(* Logix 5000 project; controller TFF vendor 1 type 14 code 107 rev 33.11; software revision 33.04; part 20 of 38 *)
(* tags used below, declared in another part *)
   Address : DINT;   // Temp Address
   Config : Configuration;   // Index Array used in configuration routines
   Index : DINT;   // Index
   TIME : DINT[2];
   TimeInSecondsDINT : DINT;
   AA008 : ALIAS FOR DigitalPoint[18];
   AI101 : ALIAS FOR AnalogPoint[16];
   AI101_SIG : ALIAS FOR DigitalPoint[106];
   AI104 : ALIAS FOR AnalogPoint[17];
   AI104_SIG : ALIAS FOR DigitalPoint[107];
   AI201A : ALIAS FOR AnalogPoint[10];
   AI201A_SIG : ALIAS FOR DigitalPoint[90];
   AI201B : ALIAS FOR AnalogPoint[0];
   AI201B_SIG : ALIAS FOR DigitalPoint[109];
   AI202 : ALIAS FOR AnalogPoint[9];
   AI202_SIG : ALIAS FOR DigitalPoint[105];
   AI203 : ALIAS FOR AnalogPoint[11];
   AI203_SIG : ALIAS FOR DigitalPoint[91];
   AI204 : ALIAS FOR AnalogPoint[12];
   AI204_SIG : ALIAS FOR DigitalPoint[92];
   AlarmAnalog : AlarmAnalog[50];   // Analog Alarm Array
   AlarmControl : AlarmControl;   // Alarm Control
   AlarmDeviation : AlarmDeviation[20];   // Control Loop Deviation Alarm Array
   AnalogOutput : AnalogOutput[25];   // Analog Output Array
   AnalogPoint : AnalogInput[50];   // Analog Input Array
   ARC_AI101 : ARC_pH;
   ARC_AI202 : ARC_pH;
   Concentration : Concentration;
   ControlLoop : ControlLoop[20];   // Control Loop Array
   ControlLoop_FeedBagLevel : ALIAS FOR ControlLoop[2];
   DF24VDC : ALIAS FOR DigitalPoint[4];
   DF24VDCPC : ALIAS FOR DigitalPoint[25];
   DF3PHP003 : ALIAS FOR DigitalPoint[27];
   DF48MIX : ALIAS FOR DigitalPoint[26];
   DF48P001 : ALIAS FOR DigitalPoint[23];
   DF48P002 : ALIAS FOR DigitalPoint[24];
   Diafiltration : Diafiltration;
   DigitalOutput : BOOL[256];   // Digital Output Array these bits are sent to output cards.
   DP : ALIAS FOR AnalogPoint[40];
   ES001 : ALIAS FOR DigitalPoint[2];
   ExternalTCU : BOOL;   // Use of External TCU
   ExternalWeight : BOOL;   // Use of External Weight
   FI003 : ALIAS FOR AnalogPoint[42];
   FI101 : ALIAS FOR AnalogPoint[19];
   FI101_SIG : ALIAS FOR DigitalPoint[110];
   FI201 : ALIAS FOR AnalogPoint[2];
   FI201_SIG : ALIAS FOR DigitalPoint[93];
   FI401 : ALIAS FOR AnalogPoint[20];
   FI401_SIG : ALIAS FOR DigitalPoint[94];
   LI101 : ALIAS FOR AnalogPoint[44];
   LI101Alarm : ALIAS FOR AlarmAnalog[44];
   MIX101 : ALIAS FOR AnalogPoint[14];
   MIX101_SIG : ALIAS FOR DigitalPoint[104];
   MIX101DF : ALIAS FOR DigitalPoint[28];
   Mixer : Mixer;   // Mixer config. structure
   NWP : ALIAS FOR AnalogPoint[45];
   Options : Options;   // Options List
   PCV101 : ALIAS FOR AnalogPoint[3];
   PCV101_Control : PCV_Control;   // PCV101 Control UDT
   PCV101_SIG : ALIAS FOR DigitalPoint[102];
   PCV201 : ALIAS FOR AnalogPoint[4];
   PCV201_Control : PCV_Control;   // PCV201 Control UDT
   PCV201_SIG : ALIAS FOR DigitalPoint[103];
   PERM : ALIAS FOR AnalogPoint[46];
   PI001 : ALIAS FOR AnalogPoint[5];
   PI001_SIG : ALIAS FOR DigitalPoint[97];
   PI101 : ALIAS FOR AnalogPoint[6];
   PI101_SIG : ALIAS FOR DigitalPoint[98];
   PI201 : ALIAS FOR AnalogPoint[7];
   PI201_SIG : ALIAS FOR DigitalPoint[99];
   PI401 : ALIAS FOR AnalogPoint[8];
   PI401_SIG : ALIAS FOR DigitalPoint[100];
   PI601 : ALIAS FOR AnalogPoint[21];
   PI601_SIG : ALIAS FOR DigitalPoint[95];
   PISL601 : ALIAS FOR DigitalPoint[0];
   PISL602 : ALIAS FOR DigitalPoint[1];
   PSH001 : ALIAS FOR DigitalPoint[21];
   PSH401 : ALIAS FOR DigitalPoint[22];
   SIC001 : ALIAS FOR Drive[1];
   SIC001DF : ALIAS FOR DigitalPoint[16];
   SIC002 : ALIAS FOR Drive[2];
   SIC002DF : ALIAS FOR DigitalPoint[17];
   SIC003DF : ALIAS FOR DigitalPoint[29];
   SIC004 : ALIAS FOR Drive[3];
   Tank : TankManagement;   // Tank Management
   TCU101 : ALIAS FOR AnalogPoint[18];
   TCU101_AO : ALIAS FOR AnalogOutput[6];
   TCU101_SIG : ALIAS FOR DigitalPoint[108];
   TCU101DF : ALIAS FOR DigitalPoint[30];
   TI101 : ALIAS FOR AnalogPoint[13];
   TI101_SIG : ALIAS FOR DigitalPoint[101];
   TI201 : ALIAS FOR AnalogPoint[22];
   TI201_SIG : ALIAS FOR DigitalPoint[111];
   TMP : ALIAS FOR AnalogPoint[41];
   Totalizer : Totalizers[20];   // Totalizers Array
   UserCr1 : ALIAS FOR DigitalPoint[65];
   UserCr2 : ALIAS FOR DigitalPoint[67];
   UserNCr1 : ALIAS FOR DigitalPoint[64];
   UserNCr2 : ALIAS FOR DigitalPoint[66];
   Valve : Valve[100];   // Valve Array
   WI101 : ALIAS FOR AnalogPoint[15];
   WI101Alarm : ALIAS FOR AlarmAnalog[15];
   WI201 : ALIAS FOR AnalogPoint[1];
   WI201_SIG : ALIAS FOR DigitalPoint[96];
   XV003 : ALIAS FOR Valve[2];
   XV004 : ALIAS FOR Valve[3];
   XV005 : ALIAS FOR Valve[4];
   XV006 : ALIAS FOR Valve[5];
   XV007 : ALIAS FOR Valve[6];
   YA01 : ALIAS FOR DigitalPoint[50];
   YA02 : ALIAS FOR DigitalPoint[51];
   YA03 : ALIAS FOR DigitalPoint[52];
   YA04 : ALIAS FOR DigitalPoint[53];
   YA05 : ALIAS FOR DigitalPoint[54];
   YA06 : ALIAS FOR DigitalPoint[55];
   YA07 : ALIAS FOR DigitalPoint[56];
   YA08 : ALIAS FOR DigitalPoint[57];
   YA09 : ALIAS FOR DigitalPoint[58];
   YA10 : ALIAS FOR DigitalPoint[59];
   YA11 : ALIAS FOR DigitalPoint[60];
   YA12 : ALIAS FOR DigitalPoint[61];
   YA13 : ALIAS FOR DigitalPoint[62];
   YA14 : ALIAS FOR DigitalPoint[63];
   YA15 : ALIAS FOR DigitalPoint[69];
   YA16 : ALIAS FOR DigitalPoint[70];
   YA17 : ALIAS FOR DigitalPoint[71];
   YA18 : ALIAS FOR DigitalPoint[72];
   YA41 : ALIAS FOR DigitalPoint[73];
   ZS008 : ALIAS FOR DigitalPoint[5];
   ZSDF : ALIAS FOR DigitalPoint[68];
(* Process, continued *)

ROUTINE Alarm_Init_Config   (* structured text *)
   (* =======================================================================
   	Alarm_Init_Config : initialize alarms to default values
   
   	List of treatments
   		- Analog alarms set point with scale Min and Max
   		- Deviation alarms
   		- Digital alarms
   	-----------------------------------------------------------------------------------------------------------------------------------------------------
   	History
   		2021-NOV-17 - Merck - Q.Spindler- Initial version for Candidate Release 1.01.00.00.a
   		2022-SEP-22 - Actemium - J. Jaekel - Modifications for Candidate Release 1.01.00.01.a
   			- Add TI201_SIG
   =============================================================================================================================*)
   
   (*Analog Set point to min/max scale, Enable alarm, timer to  2s
   ============================================================*)
   FOR Index := 0 to 49 by 1 do
   	IF AnalogPoint[Index].EnableCfg THEN
   		AlarmAnalog[Index].Override := 0; // Enable
   		AlarmAnalog[Index].LOLO := AnalogPoint[Index].ScaledMin ;
   		AlarmAnalog[Index].LO := AnalogPoint[Index].ScaledMin ;
   		AlarmAnalog[Index].HI := AnalogPoint[Index].ScaledMax ;
   		AlarmAnalog[Index].HIHI := AnalogPoint[Index].ScaledMax ;
   		AlarmAnalog[Index].LOLOTimerSP := 2 ;
   		AlarmAnalog[Index].LOTimerSP := 2 ;
   		AlarmAnalog[Index].HITimerSP := 2 ;
   		AlarmAnalog[Index].HIHITimerSP := 2 ;
   	END_IF;
   End_for ;
   
   (*Specific case for WI101
   ============================================================*)
   WI101Alarm.HI := Tank.Config.TankSelectPLC *1.2;
   WI101Alarm.HIHI := Tank.Config.TankSelectPLC *1.2;
   
   (*Specific case for LI101
   ============================================================*)
   LI101Alarm.HI := Tank.Config.TankSelectPLC;
   LI101Alarm.HIHI := Tank.Config.TankSelectPLC;
   
   (*Deviation alarm HI 100% HIHI 100%, Disable alarm, timer to 2s
   ============================================================*)
   FOR Index := 0 to 19 by 1 do
   	IF AlarmDeviation[Index].EnableCfg THEN
   		AlarmDeviation[Index].Override := 1; // Disable
   		AlarmDeviation[Index].HI := 100 ;
   		AlarmDeviation[Index].HIHI := 100 ;
   		AlarmDeviation[Index].HITimerSP := 2 ;
   		AlarmDeviation[Index].HIHITImerSP := 2 ;
   	END_IF;
   End_for ;
   
   (*Analog Set point to Disable alarm
   ============================================================*)
   // N/A
   
   (* Discrete Alarms
   ============================================================*)
   ES001.DelayTimerSP := 0;
   PISL601.Override := 0; PISL601.Priority := 1; PISL601.DelayTimerSP := 2;
   PISL602.Override := 0; PISL602.Priority := 1; PISL602.DelayTimerSP := 2;
   DF24VDC.Override := 0; DF24VDC.Priority := 1; DF24VDC.DelayTimerSP := 1;
   DF24VDCPC.Override := 0; DF24VDCPC.Priority := 1; DF24VDCPC.DelayTimerSP := 1;
   PSH001.Override := 0; PSH001.DelayTimerSP := 0;
   PSH401.Override := 0; PSH401.DelayTimerSP := 0;
   SIC001DF.Override := 0; SIC001DF.Priority := 1; SIC001DF.DelayTimerSP := 1;
   SIC002DF.Override := 0; SIC002DF.Priority := 1; SIC002DF.DelayTimerSP := 1;
   SIC003DF.Override := 0; SIC003DF.Priority := 1; SIC003DF.DelayTimerSP := 1;
   DF48P001.Override := 0; DF48P001.Priority := 1; DF48P001.DelayTimerSP := 1;
   DF48P002.Override := 0; DF48P002.Priority := 1; DF48P002.DelayTimerSP := 1;
   DF48MIX.Override := 0; DF48MIX.Priority := 1; DF48MIX.DelayTimerSP := 1;
   DF3PHP003.Override := 0; DF3PHP003.Priority := 1; DF3PHP003.DelayTimerSP := 1;
   AA008.Override := 0; AA008.Priority := 1; AA008.DelayTimerSP := 1;
   TCU101DF.Override := 0; TCU101DF.Priority := 1; TCU101DF.DelayTimerSP := 1;
   MIX101DF.Override := 0; MIX101DF.Priority := 1; MIX101DF.DelayTimerSP := 1;
   ZS008.Override := 0; ZS008.Priority := 1; ZS008.DelayTimerSP := 1;
   ZSDF.Override := 0; ZSDF.Priority := 1; ZSDF.DelayTimerSP := 1;
   
   
   YA01.Override := 0; YA01.Priority := 0; YA01.DelayTimerSP := 60;
   YA02.Override := 0; YA02.Priority := 0; YA02.DelayTimerSP := 60;
   YA03.Override := 0; YA03.Priority := 0; YA03.DelayTimerSP := 80;
   YA04.Override := 0; YA04.Priority := 0; YA04.DelayTimerSP := 60;
   YA05.Override := 0; YA05.Priority := 0; YA05.DelayTimerSP := 60;
   YA06.Override := 0; YA06.Priority := 1; YA06.DelayTimerSP := 5;
   YA07.Override := 0; YA07.Priority := 0; YA07.DelayTimerSP := 2;
   YA08.Override := 0; YA08.Priority := 1; YA08.DelayTimerSP := 5;
   YA09.Override := 0; YA09.Priority := 0; YA09.DelayTimerSP := 2;
   YA10.DelayTimerSP := 0;
   YA11.Override := 1; YA11.Priority := 0; YA11.DelayTimerSP := 5;
   YA12.Override := 0; YA12.Priority := 0; YA12.DelayTimerSP := 0;
   YA13.Override := 0; YA13.Priority := 0; YA13.DelayTimerSP := 2;
   YA14.Priority := 0; YA14.DelayTimerSP := 60;
   YA15.Override := 0; YA15.Priority := 1; YA15.DelayTimerSP := 5;
   YA16.Override := 1; YA16.Priority := 0; YA16.DelayTimerSP := 5;
   YA17.Override := 1; YA17.Priority := 0; YA17.DelayTimerSP := 5;
   YA18.Override := 0; YA18.Priority := 0; YA18.DelayTimerSP := 2;
   YA41.Override := 0; YA41.DelayTimerSP := 0;
   
   
   WI201_SIG.Override := 0; WI201_SIG.Priority := 0; WI201_SIG.DelayTimerSP := 10;
   MIX101_SIG.Override := 0; MIX101_SIG.Priority := 0; MIX101_SIG.DelayTimerSP := 10;
   AI101_SIG.Override := 0; AI101_SIG.Priority := 0; AI101_SIG.DelayTimerSP := 10;
   AI104_SIG.Override := 0; AI104_SIG.Priority := 0; AI104_SIG.DelayTimerSP := 10;
   TI101_SIG.Override := 0; TI101_SIG.Priority := 0; TI101_SIG.DelayTimerSP := 10;
   TCU101_SIG.Override := 0; TCU101_SIG.Priority := 0; TCU101_SIG.DelayTimerSP := 10;
   PI001_SIG.Override := 0; PI001_SIG.Priority := 0; PI001_SIG.DelayTimerSP := 10;
   AI201A_SIG.Override := 0; AI201A_SIG.Priority := 0; AI201A_SIG.DelayTimerSP := 10;
   AI201B_SIG.Override := 0; AI201B_SIG.Priority := 0; AI201B_SIG.DelayTimerSP := 10;
   FI201_SIG.Override := 0; FI201_SIG.Priority := 0; FI201_SIG.DelayTimerSP := 10;
   PCV201_SIG.Override := 0; PCV201_SIG.Priority := 0; PCV201_SIG.DelayTimerSP := 10;
   AI202_SIG.Override := 0; AI202_SIG.Priority := 0; AI202_SIG.DelayTimerSP := 10;
   PI201_SIG.Override := 0; PI201_SIG.Priority := 0; PI201_SIG.DelayTimerSP := 10;
   AI203_SIG.Override := 0; AI203_SIG.Priority := 0; AI203_SIG.DelayTimerSP := 10;
   AI204_SIG.Override := 0; AI204_SIG.Priority := 0; AI204_SIG.DelayTimerSP := 10;
   FI101_SIG.Override := 0; FI101_SIG.Priority := 0; FI101_SIG.DelayTimerSP := 10;
   PCV101_SIG.Override := 0; PCV101_SIG.Priority := 0; PCV101_SIG.DelayTimerSP := 10;
   PI101_SIG.Override := 0; PI101_SIG.Priority := 0; PI101_SIG.DelayTimerSP := 10;
   FI401_SIG.Override := 0; FI401_SIG.Priority := 0; FI401_SIG.DelayTimerSP := 10;
   PI401_SIG.Override := 0; PI401_SIG.Priority := 0; PI401_SIG.DelayTimerSP := 10;
   PI601_SIG.Override := 0; PI601_SIG.Priority := 0; PI601_SIG.DelayTimerSP := 10;
   TI201_SIG.Override := 0; TI201_SIG.Priority := 0; TI201_SIG.DelayTimerSP := 10;
   
   
   XV003.ZSOverride := 0; XV003.Priority := 0; XV003.AlarmTimerSP := 2;
   XV004.ZSOverride := 0; XV004.Priority := 0; XV004.AlarmTimerSP := 2;
   XV005.ZSOverride := 0; XV005.Priority := 0; XV005.AlarmTimerSP := 2;
   XV006.ZSOverride := 0; XV006.Priority := 0; XV006.AlarmTimerSP := 2;
   XV007.ZSOverride := 0; XV007.Priority := 0; XV007.AlarmTimerSP := 2;
   
   
   UserNCr1.Priority := 0; UserNCr1.DelayTimerSP := 0;
   UserCr1.Priority := 1; UserCr1.DelayTimerSP := 0;
   UserNCr2.Priority := 0; UserNCr2.DelayTimerSP := 0;
   UserCr2.Priority := 1; UserCr2.DelayTimerSP := 0;
   
   // Reset Init command
   AlarmControl.InitAlarmconfig := 0;
END_ROUTINE

ROUTINE ARCSensors_pH   (* ladder *)
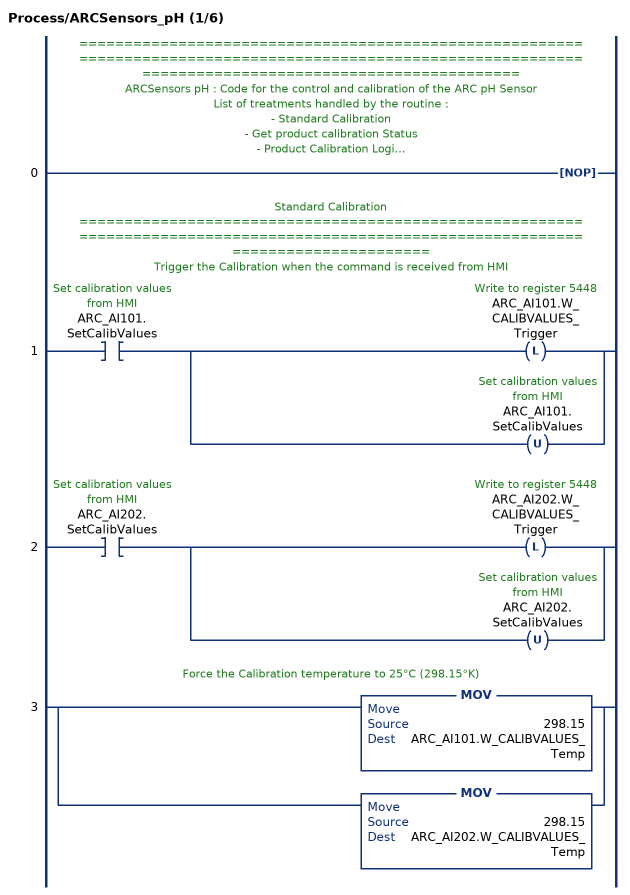
   // ==========================================================================================================================================================
   //                                                                                                                                 ARCSensors pH : Code for the control and calibration of the ARC pH Sensor
   //                                                     List of treatments handled by the routine :
   //                                             - Standard Calibration
   //                                            - Get product calibration Status
   //                                               - Product Calibration Logic
   //                                              -Set Product Calibration Commands
   //                                                     -----------------------------------------------------------------------------------------------------------------------------------------------------
   //                                                     History
   // 		2019-DEC-24 - Merck - Q. Spindler - Initial version for Candidate Release 1.00.00.00.a
   // ==========================================================================================================================================================
   0: NOP();
   // Standard Calibration
   // ======================================================================================================================================
   // Trigger the Calibration when the command is received from HMI
   1: XIC(ARC_AI101.SetCalibValues)[OTL(ARC_AI101.W_CALIBVALUES_Trigger) ,OTU(ARC_AI101.SetCalibValues) ];
   2: XIC(ARC_AI202.SetCalibValues)[OTL(ARC_AI202.W_CALIBVALUES_Trigger) ,OTU(ARC_AI202.SetCalibValues) ];
   // Force the Calibration temperature to 25°C (298.15°K)
   3: [MOV(298.15,ARC_AI101.W_CALIBVALUES_Temp) ,MOV(298.15,ARC_AI202.W_CALIBVALUES_Temp) ];
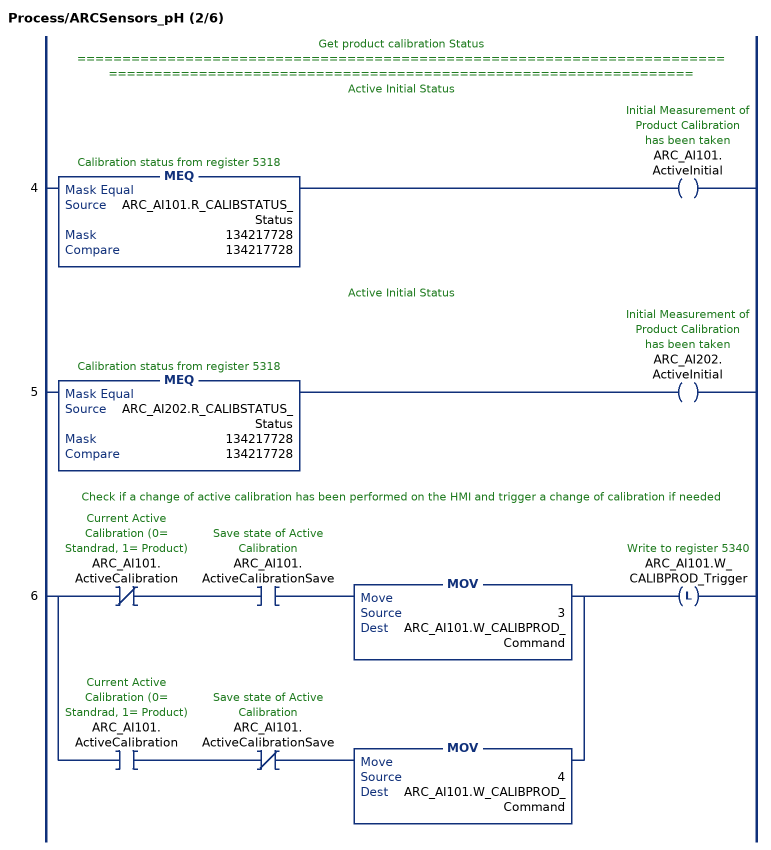
   // Get product calibration Status
   // =========================================================================================================================================
   // Active Initial Status
   4: MEQ(ARC_AI101.R_CALIBSTATUS_Status,134217728,134217728)OTE(ARC_AI101.ActiveInitial);
   // Active Initial Status
   5: MEQ(ARC_AI202.R_CALIBSTATUS_Status,134217728,134217728)OTE(ARC_AI202.ActiveInitial);
   // Check if a change of active calibration has been performed on the HMI and trigger a change of calibration if needed
   6: [XIO(ARC_AI101.ActiveCalibration) XIC(ARC_AI101.ActiveCalibrationSave) MOV(3,ARC_AI101.W_CALIBPROD_Command) ,XIC(ARC_AI101.ActiveCalibration) XIO(ARC_AI101.ActiveCalibrationSave) MOV(4,ARC_AI101.W_CALIBPROD_Command) ]OTL(ARC_AI101.W_CALIBPROD_Trigger);
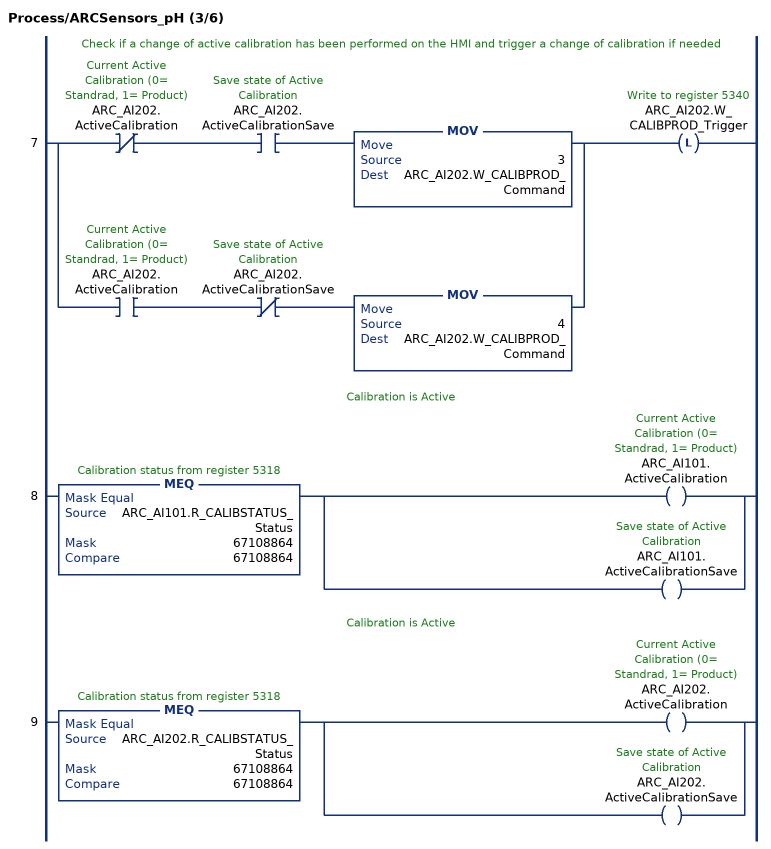
   // Check if a change of active calibration has been performed on the HMI and trigger a change of calibration if needed
   7: [XIO(ARC_AI202.ActiveCalibration) XIC(ARC_AI202.ActiveCalibrationSave) MOV(3,ARC_AI202.W_CALIBPROD_Command) ,XIC(ARC_AI202.ActiveCalibration) XIO(ARC_AI202.ActiveCalibrationSave) MOV(4,ARC_AI202.W_CALIBPROD_Command) ]OTL(ARC_AI202.W_CALIBPROD_Trigger);
   // Calibration is Active
   8: MEQ(ARC_AI101.R_CALIBSTATUS_Status,67108864,67108864)[OTE(ARC_AI101.ActiveCalibration) ,OTE(ARC_AI101.ActiveCalibrationSave) ];
   // Calibration is Active
   9: MEQ(ARC_AI202.R_CALIBSTATUS_Status,67108864,67108864)[OTE(ARC_AI202.ActiveCalibration) ,OTE(ARC_AI202.ActiveCalibrationSave) ];
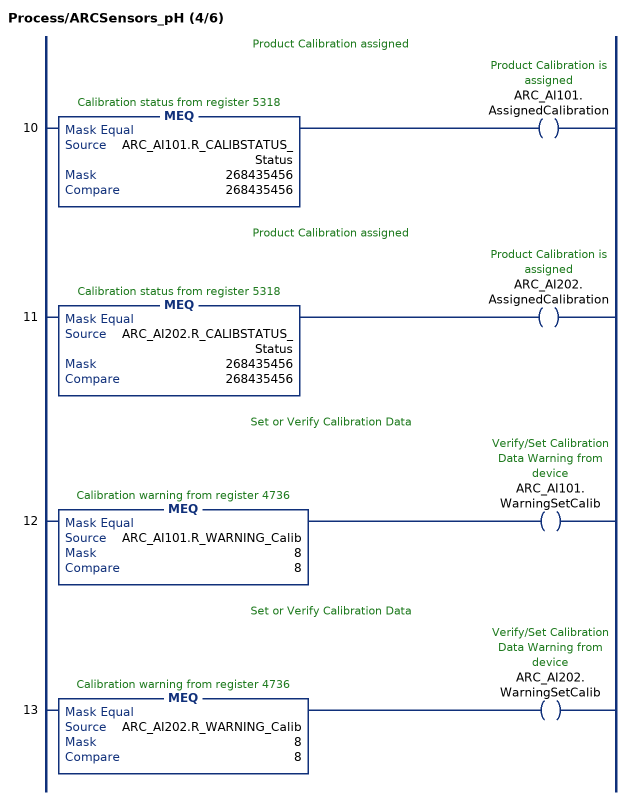
   // Product Calibration assigned
   10: MEQ(ARC_AI101.R_CALIBSTATUS_Status,268435456,268435456)OTE(ARC_AI101.AssignedCalibration);
   // Product Calibration assigned
   11: MEQ(ARC_AI202.R_CALIBSTATUS_Status,268435456,268435456)OTE(ARC_AI202.AssignedCalibration);
   // Set or Verify Calibration Data
   12: MEQ(ARC_AI101.R_WARNING_Calib,8,8)OTE(ARC_AI101.WarningSetCalib);
   // Set or Verify Calibration Data
   13: MEQ(ARC_AI202.R_WARNING_Calib,8,8)OTE(ARC_AI202.WarningSetCalib);
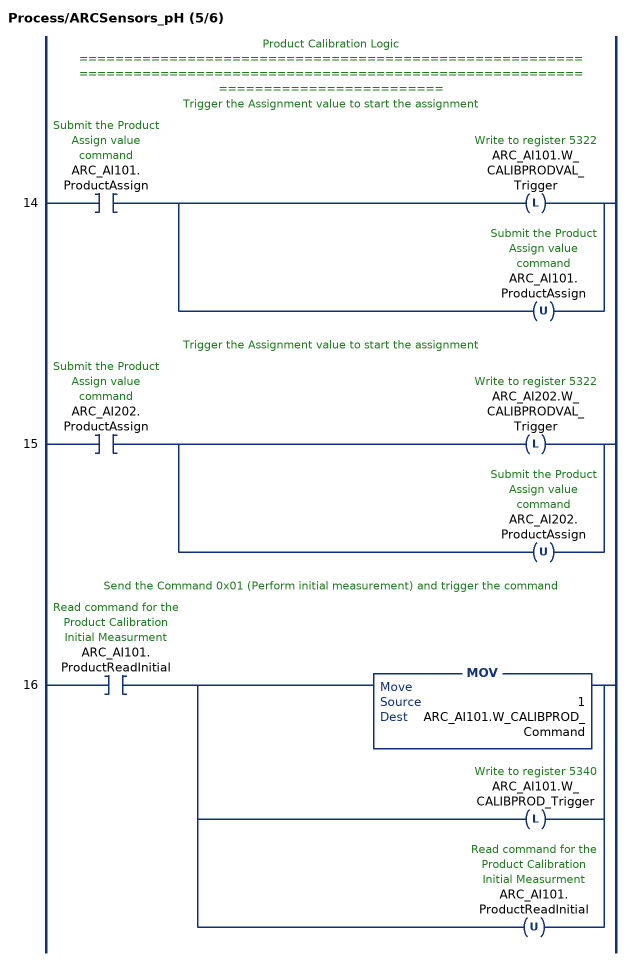
   // Product Calibration Logic
   // =========================================================================================================================================
   // Trigger the Assignment value to start the assignment
   14: XIC(ARC_AI101.ProductAssign)[OTL(ARC_AI101.W_CALIBPRODVAL_Trigger) ,OTU(ARC_AI101.ProductAssign) ];
   // Trigger the Assignment value to start the assignment
   15: XIC(ARC_AI202.ProductAssign)[OTL(ARC_AI202.W_CALIBPRODVAL_Trigger) ,OTU(ARC_AI202.ProductAssign) ];
   // Send the Command 0x01 (Perform initial measurement) and trigger the command
   16: XIC(ARC_AI101.ProductReadInitial)[MOV(1,ARC_AI101.W_CALIBPROD_Command) ,OTL(ARC_AI101.W_CALIBPROD_Trigger) ,OTU(ARC_AI101.ProductReadInitial) ];
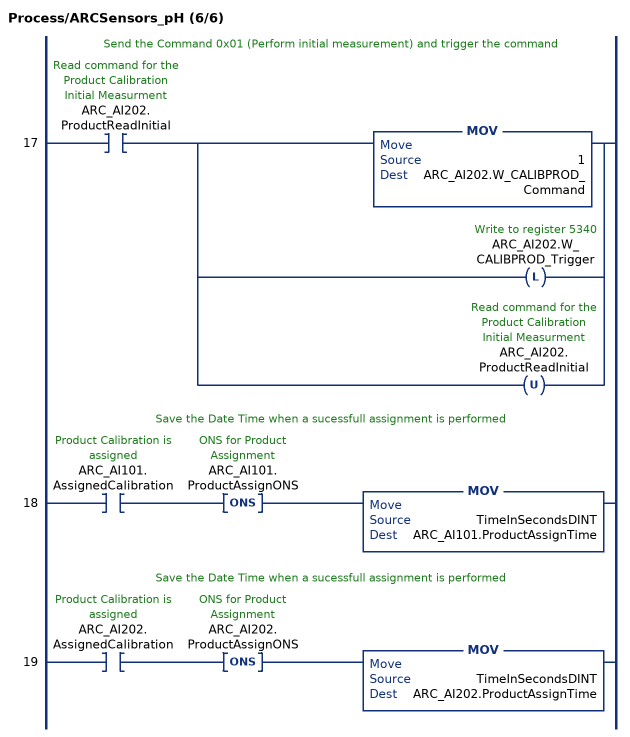
   // Send the Command 0x01 (Perform initial measurement) and trigger the command
   17: XIC(ARC_AI202.ProductReadInitial)[MOV(1,ARC_AI202.W_CALIBPROD_Command) ,OTL(ARC_AI202.W_CALIBPROD_Trigger) ,OTU(ARC_AI202.ProductReadInitial) ];
   // Save the Date Time when a sucessfull assignment is performed
   18: XIC(ARC_AI101.AssignedCalibration)ONS(ARC_AI101.ProductAssignONS)MOV(TimeInSecondsDINT,ARC_AI101.ProductAssignTime);
   // Save the Date Time when a sucessfull assignment is performed
   19: XIC(ARC_AI202.AssignedCalibration)ONS(ARC_AI202.ProductAssignONS)MOV(TimeInSecondsDINT,ARC_AI202.ProductAssignTime);
END_ROUTINE

ROUTINE Concentration_Diafiltration   (* ladder *)
// Agitator Control Routine
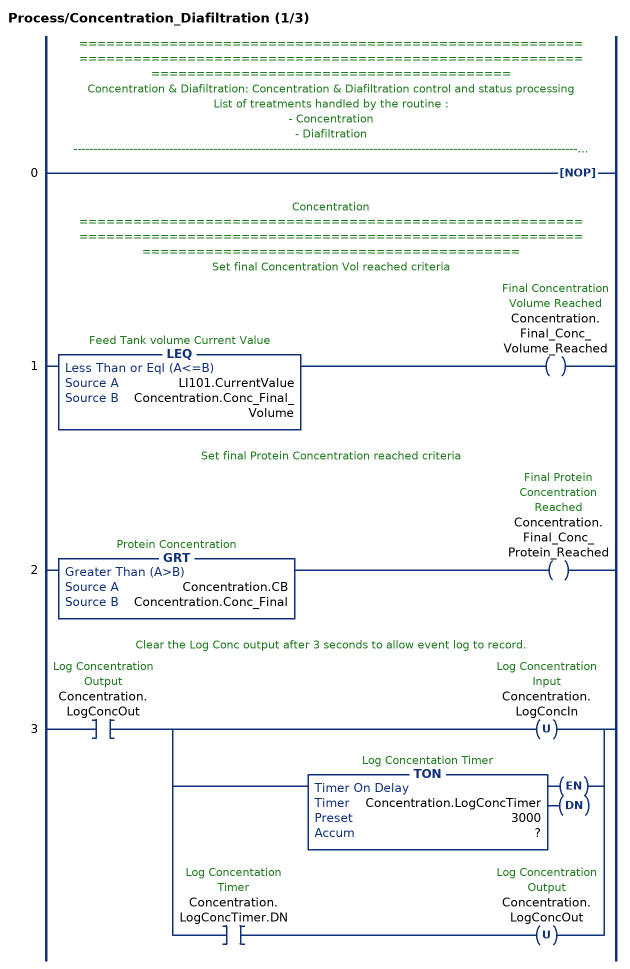
   // ========================================================================================================================================================
   //                                                                                                    Concentration & Diafiltration: Concentration & Diafiltration control and status processing
   //                                                     List of treatments handled by the routine :
   //                                                          - Concentration
   //                                                          - Diafiltration
   //                                                     -----------------------------------------------------------------------------------------------------------------------------------------------------
   //                                                     History
   // 		2019-DEC-24 - Merck - Q. Spindler - Initial version for Candidate Release 1.00.00.00.a
   // ========================================================================================================================================================
   0: NOP();
   // Concentration
   // ==========================================================================================================================================================
   // Set final Concentration Vol reached criteria
   1: LEQ(LI101.CurrentValue,Concentration.Conc_Final_Volume)OTE(Concentration.Final_Conc_Volume_Reached);
   // Set final Protein Concentration reached criteria
   2: GRT(Concentration.CB,Concentration.Conc_Final)OTE(Concentration.Final_Conc_Protein_Reached);
   // Clear the Log Conc output after 3 seconds to allow event log to record.
   3: XIC(Concentration.LogConcOut)[OTU(Concentration.LogConcIn) ,TON(Concentration.LogConcTimer,?,?) ,XIC(Concentration.LogConcTimer.DN) OTU(Concentration.LogConcOut) ];
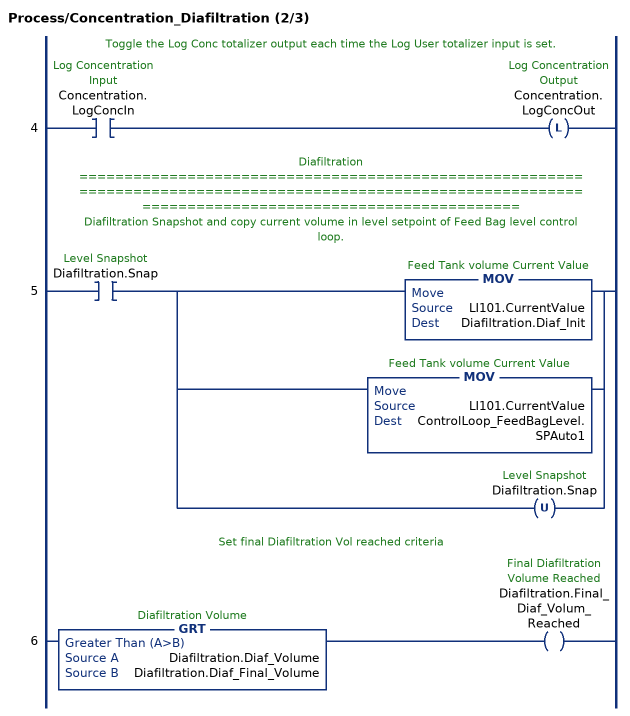
   // Toggle the Log Conc totalizer output each time the Log User totalizer input is set.
   4: XIC(Concentration.LogConcIn)OTL(Concentration.LogConcOut);
   // Diafiltration
   // ==========================================================================================================================================================
   // Diafiltration Snapshot and copy current volume in level setpoint of Feed Bag level control loop.
   5: XIC(Diafiltration.Snap)[MOV(LI101.CurrentValue,Diafiltration.Diaf_Init) ,MOV(LI101.CurrentValue,ControlLoop_FeedBagLevel.SPAuto1) ,OTU(Diafiltration.Snap) ];
   // Set final Diafiltration Vol reached criteria
   6: GRT(Diafiltration.Diaf_Volume,Diafiltration.Diaf_Final_Volume)OTE(Diafiltration.Final_Diaf_Volum_Reached);
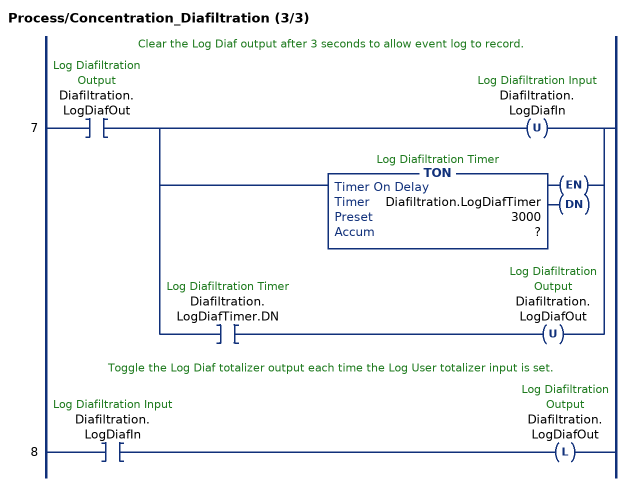
   // Clear the Log Diaf output after 3 seconds to allow event log to record.
   7: XIC(Diafiltration.LogDiafOut)[OTU(Diafiltration.LogDiafIn) ,TON(Diafiltration.LogDiafTimer,?,?) ,XIC(Diafiltration.LogDiafTimer.DN) OTU(Diafiltration.LogDiafOut) ];
   // Toggle the Log Diaf totalizer output each time the Log User totalizer input is set.
   8: XIC(Diafiltration.LogDiafIn)OTL(Diafiltration.LogDiafOut);
END_ROUTINE

ROUTINE Config_AnalogOutput   (* structured text *)
   (* ==========================================================
   	Config AnalogOutput : Configure AnalogOutput Structure
   
   	List of treatments
   		- AnalogOutput[0] : Pump P001 Speed	SIC001
   		- AnalogOutput[1] : Pump P002 Speed	SIC002
   		- AnalogOutput[2] : Pump P003 Speed	SIC003
   		- AnalogOutput[3] : PCV101 Position
   		- AnalogOutput[4] : PCV201 Position
   		- AnalogOutput[5] : Mixer MIX101 Speed SIC004
   		- AnalogOutput[6] : TCU Temperature TCU101
   		- AnalogOutput[7] : Spare AO
   		- AnalogOutput[8] : Exchange AO#1
   		- AnalogOutput[9] : Exchange AO#2
   		- AnalogOutput[10]: Exchange AO#3
   		- AnalogOutput[11]: Exchange AO#4
   		- Reset Loop : Set to 0 the AnalogOutput[12 to 24].EnableCfg
   
   -----------------------------------------------------------------------------------------------------------------------------------------------------
   	History
   		2019-DEC-24 - Merck - Q. Spindler - Initial version for Candidate Release 1.00.00.00.a
   		2021-JUN-16 - Merck - Q. Spindler - Modifications for Candidate Release 1.00.00.00.e
   					- Change TCU101 scale max to 50
   ============================================================*)
   
   (*AnalogOutput[0] : Pump P001 Speed	SIC001
   ============================================================*)
   AnalogOutput[0].EnableCfg := 1 ;
   AnalogOutput[0].RawMin := 0 ;
   AnalogOutput[0].RawMax := 27648 ;
   AnalogOutput[0].ScaledMin := 0 ;
   AnalogOutput[0].ScaledMax := 100 ;
   
   (*AnalogOutput[1] : Pump P002 Speed	SIC002
   ============================================================*)
   AnalogOutput[1].EnableCfg := 1 ;
   AnalogOutput[1].RawMin := 0 ;
   AnalogOutput[1].RawMax := 27648 ;
   AnalogOutput[1].ScaledMin := 0 ;
   AnalogOutput[1].ScaledMax := 100 ;
   
   (*AnalogOutput[2] : Pump P003 Speed	SIC003
   ============================================================*)
   AnalogOutput[2].EnableCfg := 1 ;
   AnalogOutput[2].RawMin := 0 ;
   AnalogOutput[2].RawMax := 2047 ;
   AnalogOutput[2].ScaledMin := 0 ;
   AnalogOutput[2].ScaledMax := 100 ;
   
   (*AnalogOutput[3] : PCV101 Position
   ============================================================*)
   AnalogOutput[3].EnableCfg := 1 ;
   AnalogOutput[3].RawMin := 0 ;
   AnalogOutput[3].RawMax := 2047 ;
   AnalogOutput[3].ScaledMin := 0 ;
   AnalogOutput[3].ScaledMax := 100 ;
   
   (*AnalogOutput[4] : PCV201 Position
   ============================================================*)
   AnalogOutput[4].EnableCfg := 1 ;
   AnalogOutput[4].RawMin := 0 ;
   AnalogOutput[4].RawMax := 2047 ;
   AnalogOutput[4].ScaledMin := 0 ;
   AnalogOutput[4].ScaledMax := 100 ;
   
   (*AnalogOutput[5] : Mixer MIX101 Speed SIC004
   ============================================================*)
   If Options.FeedTank then
   	AnalogOutput[5].EnableCfg := 1 ;
   else
   	AnalogOutput[5].EnableCfg := 0 ;
   End_if ;
   AnalogOutput[5].RawMin := 0 ;
   AnalogOutput[5].RawMax := 27648 ;
   AnalogOutput[5].ScaledMin := 0 ;
   AnalogOutput[5].ScaledMax := 100 ;
   
   (*AnalogOutput[6] : TCU Temperature TCU101
   ============================================================*)
   If Options.FeedTank then
   	AnalogOutput[6].EnableCfg := 1 ;
   else
   	AnalogOutput[6].EnableCfg := 0 ;
   End_if ;
   AnalogOutput[6].RawMin := 0 ;
   AnalogOutput[6].RawMax := 27648 ;
   AnalogOutput[6].ScaledMin := 0 ;
   AnalogOutput[6].ScaledMax := 50 ;
   
   (*AnalogOutput[7] : Spare AO
   ============================================================*)
   AnalogOutput[7].EnableCfg := 0 ;
   AnalogOutput[7].RawMin := 0 ;
   AnalogOutput[7].RawMax := 27648 ;
   AnalogOutput[7].ScaledMin := 0 ;
   AnalogOutput[7].ScaledMax := 100 ;
   
   (*AnalogOutput[8] : Exchange AO#1
   ============================================================*)
   (*Set to 1 to use this AnalogOut*)
   If Options.External_IO then
   	AnalogOutput[8].EnableCfg := 1 ;
   else
   	AnalogOutput[8].EnableCfg := 0 ;
   End_if ;
   (*Default Configuration *)
   AnalogOutput[8].RawMin := 0 ;
   AnalogOutput[8].RawMax := 2047 ;
   AnalogOutput[8].ScaledMin := 0 ;
   AnalogOutput[8].ScaledMax := 100 ;
   
   (*AnalogOutput[9] : Exchange AO#2
   ============================================================*)
   (*Set to 1 to use this AnalogOut*)
   If Options.External_IO then
   	AnalogOutput[9].EnableCfg := 1 ;
   else
   	AnalogOutput[9].EnableCfg := 0 ;
   End_if ;
   (*Default Configuration *)
   AnalogOutput[9].RawMin := 0 ;
   AnalogOutput[9].RawMax := 2047 ;
   AnalogOutput[9].ScaledMin := 0 ;
   AnalogOutput[9].ScaledMax := 100 ;
   
   (*AnalogOutput[10]: Exchange AO#3
   ============================================================*)
   (*Set to 1 to use this AnalogOut*)
   If Options.External_IO then
   	AnalogOutput[10].EnableCfg := 1 ;
   else
   	AnalogOutput[10].EnableCfg := 0 ;
   End_if ;
   (*Default Configuration *)
   AnalogOutput[10].RawMin := 0 ;
   AnalogOutput[10].RawMax := 2047 ;
   AnalogOutput[10].ScaledMin := 0 ;
   AnalogOutput[10].ScaledMax := 100 ;
   
   (*AnalogOutput[11]: Exchange AO#4
   ============================================================*)
   (*Set to 1 to use this AnalogOut*)
   If Options.External_IO then
   	AnalogOutput[11].EnableCfg := 1 ;
   else
   	AnalogOutput[11].EnableCfg := 0 ;
   End_if ;
   (*Default Configuration *)
   AnalogOutput[11].RawMin := 0 ;
   AnalogOutput[11].RawMax := 2047 ;
   AnalogOutput[11].ScaledMin := 0 ;
   AnalogOutput[11].ScaledMax := 100 ;
   
   (*Reset Loop : Set to 0 the AnalogOutput[12 to 24].EnableCfg
   ============================================================*)
   FOR Config.IndexA0 := 5 to 24 by 1 do
   	AnalogOutput[Config.IndexA0].EnableCfg := 0 ;
   End_for ;
   
END_ROUTINE

ROUTINE Config_AnalogPoint   (* structured text *)
// Apply the default configuration
   (* ==========================================================
   	Config AnalogPoint : Configure AnalogPoint Structure
   
   	List of treatments
   		- AnalogPoint[0] : Filtrate Conductivity Cleaning AI201B
   		- AnalogPoint[1] : External Filtrate Weight Scale WI201
   		- AnalogPoint[2] : Filtrate Flow FI201
   		- AnalogPoint[3] : Retentate Pressure Control Valve Position PCV101
   		- AnalogPoint[4] : Filtrate Pressure Control Valve Position PCV201
   		- AnalogPoint[5] : Feed Pressure PI001
   		- AnalogPoint[6] : Retentate Pressure PI101
   		- AnalogPoint[7] : Filtrate Pressure PI201
   		- AnalogPoint[8] : Transfer Pump Pressure PI401
   		- AnalogPoint[9] : Filtrate pH AI202
   		- AnalogPoint[10]: Filtrate Conductivity Process AI201A
   		- AnalogPoint[11]: Filtrate UV AI203
   		- AnalogPoint[12]: Filtrate UV AI204
   		- AnalogPoint[13]: Feed Tank Temperature TI101
   		- AnalogPoint[14]: Mixer Speed MIX101
   		- AnalogPoint[15]: Feed Tank Weight WI101
   		- AnalogPoint[16]: Feed Tank pH AI101
   		- AnalogPoint[17]: Feed Tank Conductivity AI104
   		- AnalogPoint[18]: TCU Temperature TCU101
   		- AnalogPoint[19]: Retentate Flow FI101
   		- AnalogPoint[20]: Transfer Pump Flow FI401
   		- AnalogPoint[21]: Feed Tank Pressure PI601
   		- AnalogPoint[22]: Filtrate Temperature TI201
   		- Reset Loop : Set to 0 the AnalogPoint[23 to 27].EnableCfg
   		- AnalogPoint[28]: Exchange AI#1
   		- AnalogPoint[29]: Exchange AI#2
   		- AnalogPoint[30]: Exchange AI#3
   		- AnalogPoint[31]: Exchange AI#4
   		- Reset Loop : Set to 0 the AnalogPoint[32 to 39].EnableCfg
   		- AnalogPoint[40]: Differential Pressure DP
   		- AnalogPoint[41]: Trans-Membrane Pressure TMP
   		- AnalogPoint[42]: Feed Flow FI003
   		- AnalogPoint[43]: Spare
   		- AnalogPoint[44]: Feed Tank Volume LI101
   		- AnalogPoint[45]: Normalized Water Permeability NWP
   		- AnalogPoint[46]: Membrane Permeability PERM
   		- Reset Loop : Set to 0 the AnalogPoint[47 to 49].EnableCfg
   
   -----------------------------------------------------------------------------------------------------------------------------------------------------
   	History
   		2019-DEC-24 - Merck - Q. Spindler - Initial version for Candidate Release 1.00.00.00.a
   		2020-MAR-25 - Merck - Q. Spindler - Modifications for Candidate Release 1.00.00.00.b
   					- Change MIX101 Raw Values to match 0-5V input
   					- Change MIX101, TCU101, TI101, AI104 Raw Values to match 56200 IO Card
   		2020-SEP-18 - Merck - Q. Spindler - Modifications for Candidate Release 1.00.00.00.d
   					- Disable WI201 alarm if ExternalWeight not used
   		2021-APR-15 - Merck - Q. Spindler - Modifications for Candidate Release 1.00.00.00.e
   					- Disable HIHIEnable (so HIHI Alarm are no longer forced ON) for PI001, PI101, PI201, and PI401
   					- Add FiltrateUltrasonicFlow option for FI201
   					- Add RawLowLimit to 2mA for PI001, PI101, PI201, PI401, and PI601
   		2022-SEP-22 - Actemium - J. Jaekel - Modifications for Candidate Release 1.01.00.01.a
   					- Add ExternalTCU option to TCU101 AnalogPoint
   					- Add AnalogPoint[22]: Filtrate Temperature TI201
   		2022-NOV-21 - Actemium - J. Jaekel - Modifications for Candidate Release 1.01.00.01.b
   					- Update of TI201 enable condition
   ============================================================*)
   
   
   (*AnalogPoint[0] : Filtrate Conductivity Cleaning AI201B
   ============================================================*)
   IF Options.FiltrateCondPHUV OR Options.FiltrateCondPH THEN
   	AnalogPoint[0].EnableCfg := 1 ;
   	AlarmAnalog[0].EnableCfg := 1 ;
   ELSE
   	AnalogPoint[0].EnableCfg := 0 ;
   	AlarmAnalog[0].EnableCfg := 0 ;
   END_IF;
   AnalogPoint[0].Address := 0 ;
   AnalogPoint[0].RawMin := 5529 ;
   AnalogPoint[0].RawMax := 27648 ;
   AnalogPoint[0].RealCfg := 1 ;
   AnalogPoint[0].OverrideCfg := 1 ;
   AlarmAnalog[0].FeedPumpEnable := 0 ;
   AlarmAnalog[0].FeedPumpTag := 0 ;
   AlarmAnalog[0].TransferPumpEnable := 0 ;
   AlarmAnalog[0].TransferPumpTag := 0 ;
   AlarmAnalog[0].Disable := 0 ;
   AlarmAnalog[0].HIHIEnable := 0 ;
   
   (*AnalogPoint[1] : External Filtrate Weight Scale WI201
   ============================================================*)
   IF ExternalWeight THEN
   	AlarmAnalog[1].EnableCfg := 1 ;
   ELSE
   	AlarmAnalog[1].EnableCfg := 0 ;
   	AlarmAnalog[1].ValueHMI := 0 ;
   	AlarmAnalog[1].LOAlarm := 0 ;
   	AlarmAnalog[1].LOLOAlarm := 0 ;
   	AlarmAnalog[1].HIAlarm := 0 ;
   	AlarmAnalog[1].HIHIAlarm := 0 ;
   END_IF;
   AnalogPoint[1].EnableCfg := 1 ;
   AnalogPoint[1].Address := 1 ;
   AnalogPoint[1].RawMin := 6553 ;
   AnalogPoint[1].RawMax := 32767 ;
   AnalogPoint[1].RealCfg := 1 ;
   AnalogPoint[1].OverrideCfg := 1 ;
   AlarmAnalog[1].FeedPumpEnable := 0 ;
   AlarmAnalog[1].FeedPumpTag := 0 ;
   AlarmAnalog[1].TransferPumpEnable := 0 ;
   AlarmAnalog[1].TransferPumpTag := 0 ;
   AlarmAnalog[1].Disable := 0 ;
   AlarmAnalog[1].HIHIEnable := 0 ;
   
   (*AnalogPoint[2] : Filtrate Flow FI201
   ============================================================*)
   AnalogPoint[2].EnableCfg := 1 ;
   AlarmAnalog[2].EnableCfg := 1 ;
   IF Options.FiltrateUltrasonicFlow THEN
   	AnalogPoint[2].RealCfg := 1 ;
   ELSE
   	AnalogPoint[2].RealCfg := 0 ; // For Qmax Factor
   END_IF;
   AnalogPoint[2].Address := 2 ;
   AnalogPoint[2].RawMin := 6553 ;
   AnalogPoint[2].RawMax := 32767 ;
   AnalogPoint[2].OverrideCfg := 1 ;
   AlarmAnalog[2].FeedPumpEnable := 1 ;
   AlarmAnalog[2].FeedPumpTag := 1 ;
   AlarmAnalog[2].TransferPumpEnable := 0 ;
   AlarmAnalog[2].TransferPumpTag := 0 ;
   AlarmAnalog[2].Disable := 0 ;
   AlarmAnalog[2].HIHIEnable := 0 ;
   
   (*AnalogPoint[3] : Retentate Pressure Control Valve Position PCV101
   ============================================================*)
   AnalogPoint[3].EnableCfg := 1 ;
   AlarmAnalog[3].EnableCfg := 0 ;
   AnalogPoint[3].Address := 3 ;
   AnalogPoint[3].RawMin := 6553 ;
   AnalogPoint[3].RawMax := 32767 ;
   AnalogPoint[3].RealCfg := 0 ;
   AnalogPoint[3].OverrideCfg := 0 ;
   AlarmAnalog[3].FeedPumpEnable := 0 ;
   AlarmAnalog[3].FeedPumpTag := 0 ;
   AlarmAnalog[3].TransferPumpEnable := 0 ;
   AlarmAnalog[3].TransferPumpTag := 0 ;
   AlarmAnalog[3].Disable := 0 ;
   AlarmAnalog[3].HIHIEnable := 0 ;
   
   (*AnalogPoint[4] : Filtrate Pressure Control Valve Position PCV201
   ============================================================*)
   AnalogPoint[4].EnableCfg := 1 ;
   AlarmAnalog[4].EnableCfg := 0 ;
   AnalogPoint[4].Address := 4 ;
   AnalogPoint[4].RawMin := 6553 ;
   AnalogPoint[4].RawMax := 32767 ;
   AnalogPoint[4].RealCfg := 0 ;
   AnalogPoint[4].OverrideCfg := 0 ;
   AlarmAnalog[4].FeedPumpEnable := 0 ;
   AlarmAnalog[4].FeedPumpTag := 0 ;
   AlarmAnalog[4].TransferPumpEnable := 0 ;
   AlarmAnalog[4].TransferPumpTag := 0 ;
   AlarmAnalog[4].Disable := 0 ;
   AlarmAnalog[4].HIHIEnable := 0 ;
   
   (*AnalogPoint[5] : Feed Pressure PI001
   ============================================================*)
   AnalogPoint[5].EnableCfg := 1 ;
   AlarmAnalog[5].EnableCfg := 1 ;
   AnalogPoint[5].Address := 5 ;
   AnalogPoint[5].RawMin := 6553 ;
   AnalogPoint[5].RawMax := 32767 ;
   AnalogPoint[5].RawLowLimit := 3276; // 2mA
   AnalogPoint[5].RealCfg := 1 ;
   AnalogPoint[5].OverrideCfg := 1 ;
   AlarmAnalog[5].FeedPumpEnable := 1 ;
   AlarmAnalog[5].FeedPumpTag := 1 ;
   AlarmAnalog[5].TransferPumpEnable := 0 ;
   AlarmAnalog[5].TransferPumpTag := 0 ;
   AlarmAnalog[5].Disable := 0 ;
   AlarmAnalog[5].HIHIEnable := 0 ;
   
   (*AnalogPoint[6] : Retentate Pressure PI101
   ============================================================*)
   AnalogPoint[6].EnableCfg := 1 ;
   AlarmAnalog[6].EnableCfg := 1 ;
   AnalogPoint[6].Address := 6 ;
   AnalogPoint[6].RawMin := 6553 ;
   AnalogPoint[6].RawMax := 32767 ;
   AnalogPoint[6].RawLowLimit := 3276; // 2mA
   AnalogPoint[6].RealCfg := 1 ;
   AnalogPoint[6].OverrideCfg := 1 ;
   AlarmAnalog[6].FeedPumpEnable := 1 ;
   AlarmAnalog[6].FeedPumpTag := 1 ;
   AlarmAnalog[6].TransferPumpEnable := 0 ;
   AlarmAnalog[6].TransferPumpTag := 0 ;
   AlarmAnalog[6].Disable := 0 ;
   AlarmAnalog[6].HIHIEnable := 0 ;
   
   (*AnalogPoint[7] : Filtrate Pressure PI201
   ============================================================*)
   AnalogPoint[7].EnableCfg := 1 ;
   AlarmAnalog[7].EnableCfg := 1 ;
   AnalogPoint[7].Address := 7 ;
   AnalogPoint[7].RawMin := 6553 ;
   AnalogPoint[7].RawMax := 32767 ;
   AnalogPoint[7].RawLowLimit := 3276; // 2mA
   AnalogPoint[7].RealCfg := 1 ;
   AnalogPoint[7].OverrideCfg := 1 ;
   AlarmAnalog[7].FeedPumpEnable := 1 ;
   AlarmAnalog[7].FeedPumpTag := 1 ;
   AlarmAnalog[7].TransferPumpEnable := 0 ;
   AlarmAnalog[7].TransferPumpTag := 0 ;
   AlarmAnalog[7].Disable := 0 ;
   AlarmAnalog[7].HIHIEnable := 0 ;
   
   (*AnalogPoint[8] : Transfer Pump Pressure PI401
   ============================================================*)
   AnalogPoint[8].EnableCfg := 1 ;
   AlarmAnalog[8].EnableCfg := 1 ;
   AnalogPoint[8].Address := 8 ;
   AnalogPoint[8].RawMin := 6553 ;
   AnalogPoint[8].RawMax := 32767 ;
   AnalogPoint[8].RawLowLimit := 3276; // 2mA
   AnalogPoint[8].RealCfg := 1 ;
   AnalogPoint[8].OverrideCfg := 1 ;
   AlarmAnalog[8].FeedPumpEnable := 0 ;
   AlarmAnalog[8].FeedPumpTag := 0 ;
   AlarmAnalog[8].TransferPumpEnable := 1 ;
   AlarmAnalog[8].TransferPumpTag := 2 ;
   AlarmAnalog[8].Disable := 0 ;
   AlarmAnalog[8].HIHIEnable := 0 ;
   
   (*AnalogPoint[9] : Filtrate pH AI202
   ============================================================*)
   IF Options.FiltrateCondPHUV OR Options.FiltrateCondPH THEN
   	AnalogPoint[9].EnableCfg := 1 ;
   	AlarmAnalog[9].EnableCfg := 1 ;
   	IF Options.SingleUsePH THEN
   		AnalogPoint[9].RealCfg := 0 ;
   	ELSE
   		AnalogPoint[9].RealCfg := 1 ;
   	END_IF;
   ELSE
   	AnalogPoint[9].EnableCfg := 0 ;
   	AlarmAnalog[9].EnableCfg := 0 ;
   	AnalogPoint[9].RealCfg := 1 ;
   END_IF;
   AnalogPoint[9].Address := 9 ;
   AnalogPoint[9].RawMin := 5529 ;
   AnalogPoint[9].RawMax := 27648 ;
   AnalogPoint[9].OverrideCfg := 1 ;
   AlarmAnalog[9].FeedPumpEnable := 0 ;
   AlarmAnalog[9].FeedPumpTag := 0 ;
   AlarmAnalog[9].TransferPumpEnable := 0 ;
   AlarmAnalog[9].TransferPumpTag := 0 ;
   AlarmAnalog[9].Disable := 0 ;
   AlarmAnalog[9].HIHIEnable := 0 ;
   
   (*AnalogPoint[10]: Filtrate Conductivity Process AI201A
   ============================================================*)
   IF Options.FiltrateCondPHUV OR Options.FiltrateCondPH THEN
   	AnalogPoint[10].EnableCfg := 1 ;
   	AlarmAnalog[10].EnableCfg := 1 ;
   ELSE
   	AnalogPoint[10].EnableCfg := 0 ;
   	AlarmAnalog[10].EnableCfg := 0 ;
   END_IF;
   AnalogPoint[10].Address := 10 ;
   AnalogPoint[10].RawMin := 5529 ;
   AnalogPoint[10].RawMax := 27648 ;
   AnalogPoint[10].RealCfg := 1 ;
   AnalogPoint[10].OverrideCfg := 1 ;
   AlarmAnalog[10].FeedPumpEnable := 0 ;
   AlarmAnalog[10].FeedPumpTag := 0 ;
   AlarmAnalog[10].TransferPumpEnable := 0 ;
   AlarmAnalog[10].TransferPumpTag := 0 ;
   AlarmAnalog[10].Disable := 0 ;
   AlarmAnalog[10].HIHIEnable := 0 ;
   
   (*AnalogPoint[11]: Filtrate UV AI203
   ============================================================*)
   IF Options.FiltrateCondPHUV THEN
   	AnalogPoint[11].EnableCfg := 1 ;
   	AlarmAnalog[11].EnableCfg := 1 ;
   ELSE
   	AnalogPoint[11].EnableCfg := 0 ;
   	AlarmAnalog[11].EnableCfg := 0 ;
   END_IF;
   AnalogPoint[11].Address := 11 ;
   AnalogPoint[11].RawMin := 5529 ;
   AnalogPoint[11].RawMax := 27648 ;
   AnalogPoint[11].RealCfg := 1 ;
   AnalogPoint[11].OverrideCfg := 1 ;
   AlarmAnalog[11].FeedPumpEnable := 0 ;
   AlarmAnalog[11].FeedPumpTag := 0 ;
   AlarmAnalog[11].TransferPumpEnable := 0 ;
   AlarmAnalog[11].TransferPumpTag := 0 ;
   AlarmAnalog[11].Disable := 0 ;
   AlarmAnalog[11].HIHIEnable := 0 ;
   
   (*AnalogPoint[12]: Filtrate UV AI204
   ============================================================*)
   IF Options.FiltrateCondPHUV THEN
   	AnalogPoint[12].EnableCfg := 1 ;
   	AlarmAnalog[12].EnableCfg := 1 ;
   ELSE
   	AnalogPoint[12].EnableCfg := 0 ;
   	AlarmAnalog[12].EnableCfg := 0 ;
   END_IF;
   AnalogPoint[12].Address := 12 ;
   AnalogPoint[12].RawMin := 5529 ;
   AnalogPoint[12].RawMax := 27648 ;
   AnalogPoint[12].RealCfg := 1 ;
   AnalogPoint[12].OverrideCfg := 1 ;
   AlarmAnalog[12].FeedPumpEnable := 0 ;
   AlarmAnalog[12].FeedPumpTag := 0 ;
   AlarmAnalog[12].TransferPumpEnable := 0 ;
   AlarmAnalog[12].TransferPumpTag := 0 ;
   AlarmAnalog[12].Disable := 0 ;
   AlarmAnalog[12].HIHIEnable := 0 ;
   
   (*AnalogPoint[13]: Feed Tank Temperature TI101
   ============================================================*)
   IF Options.FeedTank THEN
   	AnalogPoint[13].EnableCfg := 1 ;
   	AlarmAnalog[13].EnableCfg := 1 ;
   ELSE
   	AnalogPoint[13].EnableCfg := 0 ;
   	AlarmAnalog[13].EnableCfg := 0 ;
   END_IF;
   AnalogPoint[13].Address := 13 ;
   AnalogPoint[13].RawMin := 5529 ;
   AnalogPoint[13].RawMax := 27648 ;
   AnalogPoint[13].RealCfg := 1 ;
   AnalogPoint[13].OverrideCfg := 1 ;
   AlarmAnalog[13].FeedPumpEnable := 0 ;
   AlarmAnalog[13].FeedPumpTag := 0 ;
   AlarmAnalog[13].TransferPumpEnable := 0 ;
   AlarmAnalog[13].TransferPumpTag := 0 ;
   AlarmAnalog[13].Disable := 0 ;
   AlarmAnalog[13].HIHIEnable := 0 ;
   
   (*AnalogPoint[14]: Mixer Speed MIX101
   ============================================================*)
   IF Options.FeedTank THEN
   	AnalogPoint[14].EnableCfg := 1 ;
   ELSE
   	AnalogPoint[14].EnableCfg := 0 ;
   END_IF;
   AnalogPoint[14].Address := 14 ;
   AnalogPoint[14].RawMin := 0 ;
   AnalogPoint[14].RawMax := 13824 ; // 27648 / 2 to scale a 0-10V to 0-5V input
   AnalogPoint[14].RealCfg := 1 ;
   AnalogPoint[14].OverrideCfg := 0 ;
   AlarmAnalog[14].FeedPumpEnable := 0 ;
   AlarmAnalog[14].FeedPumpTag := 0 ;
   AlarmAnalog[14].TransferPumpEnable := 0 ;
   AlarmAnalog[14].TransferPumpTag := 0 ;
   AlarmAnalog[14].EnableCfg := 0 ;
   AlarmAnalog[14].Disable := 0 ;
   AlarmAnalog[14].HIHIEnable := 0 ;
   
   (*AnalogPoint[15]: Feed Tank Weight WI101
   ============================================================*)
   AnalogPoint[15].EnableCfg := 1 ;
   AlarmAnalog[15].EnableCfg := 1 ;
   AnalogPoint[15].Address := 15 ;
   AnalogPoint[15].RawMin := 0 ;
   AnalogPoint[15].RawMax := 99999 ;
   AnalogPoint[15].RealCfg := 0 ;
   AnalogPoint[15].OverrideCfg := 1 ;
   AnalogPoint[15].ScaledMin := 0 ;
   AnalogPoint[15].ScaledMax := 999.99 ;
   AlarmAnalog[15].FeedPumpEnable := 1 ;
   AlarmAnalog[15].FeedPumpTag := 1 ;
   AlarmAnalog[15].TransferPumpEnable := 0 ;
   AlarmAnalog[15].TransferPumpTag := 0 ;
   AlarmAnalog[15].Disable := 0 ;
   AlarmAnalog[15].HIHIDisable := NOT SIC002.RunStatus ;
   AlarmAnalog[15].HIDisable := NOT SIC002.RunStatus ;
   AlarmAnalog[15].HIHIEnable := 0 ;
   
   (*AnalogPoint[16]: Feed Tank pH AI101
   ============================================================*)
   IF Options.FeedTank AND Options.TankPH THEN
   	AnalogPoint[16].EnableCfg := 1 ;
   	AlarmAnalog[16].EnableCfg := 1 ;
   ELSE
   	AnalogPoint[16].EnableCfg := 0 ;
   	AlarmAnalog[16].EnableCfg := 0 ;
   END_IF;
   AnalogPoint[16].Address := 16 ;
   AnalogPoint[16].RawMin := 6553 ;
   AnalogPoint[16].RawMax := 32767 ;
   AnalogPoint[16].RealCfg := 0 ;
   AnalogPoint[16].OverrideCfg := 1 ;
   AlarmAnalog[16].FeedPumpEnable := 0 ;
   AlarmAnalog[16].FeedPumpTag := 0 ;
   AlarmAnalog[16].TransferPumpEnable := 0 ;
   AlarmAnalog[16].TransferPumpTag := 0 ;
   AlarmAnalog[16].Disable := 0 ;
   AlarmAnalog[16].HIHIEnable := 0 ;
   
   (*AnalogPoint[17]: Feed Tank Conductivity AI104
   ============================================================*)
   IF Options.FeedTank AND Options.TankCond THEN
   	AnalogPoint[17].EnableCfg := 1 ;
   	AlarmAnalog[17].EnableCfg := 1 ;
   ELSE
   	AnalogPoint[17].EnableCfg := 0 ;
   	AlarmAnalog[17].EnableCfg := 0 ;
   END_IF;
   AnalogPoint[17].Address := 17 ;
   AnalogPoint[17].RawMin := 5529 ;
   AnalogPoint[17].RawMax := 27648 ;
   AnalogPoint[17].RealCfg := 1 ;
   AnalogPoint[17].OverrideCfg := 1 ;
   AlarmAnalog[17].FeedPumpEnable := 0 ;
   AlarmAnalog[17].FeedPumpTag := 0 ;
   AlarmAnalog[17].TransferPumpEnable := 0 ;
   AlarmAnalog[17].TransferPumpTag := 0 ;
   AlarmAnalog[17].Disable := 0 ;
   AlarmAnalog[17].HIHIEnable := 0 ;
   
   (*AnalogPoint[18]: TCU Temperature TCU101
   ============================================================*)
   IF Options.FeedTank and ExternalTCU THEN
   	AnalogPoint[18].EnableCfg := 1 ;
   ELSE
   	AnalogPoint[18].EnableCfg := 0 ;
   END_IF;
   AnalogPoint[18].Address := 18 ;
   AnalogPoint[18].RawMin := 5529 ;
   AnalogPoint[18].RawMax := 27648 ;
   AnalogPoint[18].RealCfg := 1 ;
   AnalogPoint[18].OverrideCfg := 1 ;
   AlarmAnalog[18].EnableCfg := 0 ;
   AlarmAnalog[18].FeedPumpEnable := 0 ;
   AlarmAnalog[18].FeedPumpTag := 0 ;
   AlarmAnalog[18].TransferPumpEnable := 0 ;
   AlarmAnalog[18].TransferPumpTag := 0 ;
   AlarmAnalog[18].Disable := 0 ;
   AlarmAnalog[18].HIHIEnable := 0 ;
   
   (*AnalogPoint[19]: Retentate Flow FI101
   ============================================================*)
   AnalogPoint[19].EnableCfg := 1 ;
   AlarmAnalog[19].EnableCfg := 1 ;
   AnalogPoint[19].Address := 19 ;
   AnalogPoint[19].RawMin := 6553 ;
   AnalogPoint[19].RawMax := 32767 ;
   AnalogPoint[19].RealCfg := 0 ; // For Qmax Factor
   AnalogPoint[19].OverrideCfg := 1 ;
   AlarmAnalog[19].FeedPumpEnable := 1 ;
   AlarmAnalog[19].FeedPumpTag := 1 ;
   AlarmAnalog[19].TransferPumpEnable := 0 ;
   AlarmAnalog[19].TransferPumpTag := 0 ;
   AlarmAnalog[19].Disable := 0 ;
   AlarmAnalog[19].HIHIEnable := 0 ;
   
   (*AnalogPoint[20]: Transfer Pump Flow FI401
   ============================================================*)
   IF Options.TransferFlow THEN
   	AnalogPoint[20].EnableCfg := 1 ;
   	AlarmAnalog[20].EnableCfg := 1 ;
   ELSE
   	AnalogPoint[20].EnableCfg := 0 ;
   	AlarmAnalog[20].EnableCfg := 0 ;
   END_IF;
   AnalogPoint[20].Address := 20 ;
   AnalogPoint[20].RawMin := 6553 ;
   AnalogPoint[20].RawMax := 32767 ;
   AnalogPoint[20].RealCfg := 0 ; // For Qmax Factor
   AnalogPoint[20].OverrideCfg := 1 ;
   AlarmAnalog[20].FeedPumpEnable := 0 ;
   AlarmAnalog[20].FeedPumpTag := 0 ;
   AlarmAnalog[20].TransferPumpEnable := 1 ;
   AlarmAnalog[20].TransferPumpTag := 2 ;
   AlarmAnalog[20].Disable := 0 ;
   AlarmAnalog[20].HIHIEnable := 0 ;
   
   (*AnalogPoint[21]: Feed Tank Pressure PI601
   ============================================================*)
   IF Options.FeedTank THEN
   	AnalogPoint[21].EnableCfg := 1 ;
   	AlarmAnalog[21].EnableCfg := 1 ;
   ELSE
   	AnalogPoint[21].EnableCfg := 0 ;
   	AlarmAnalog[21].EnableCfg := 0 ;
   END_IF;
   AnalogPoint[21].Address := 21 ;
   AnalogPoint[21].RawMin := 6553 ;
   AnalogPoint[21].RawMax := 32767 ;
   AnalogPoint[21].RawLowLimit := 3276; // 2mA
   AnalogPoint[21].RealCfg := 1 ;
   AnalogPoint[21].OverrideCfg := 1 ;
   AlarmAnalog[21].FeedPumpEnable := 0 ;
   AlarmAnalog[21].FeedPumpTag := 0 ;
   AlarmAnalog[21].TransferPumpEnable := 0 ;
   AlarmAnalog[21].TransferPumpTag := 0 ;
   AlarmAnalog[21].Disable := 0 ;
   AlarmAnalog[21].HIHIEnable := 0 ;
   
   (*AnalogPoint[22] : Filtrate Temperature TI201
   ============================================================*)
   IF Options.FiltrateCondPHUV OR Options.FiltrateCondPH THEN
   	AnalogPoint[22].EnableCfg := 1 ;
   	AlarmAnalog[22].EnableCfg := 1 ;
   ELSE
   	AnalogPoint[22].EnableCfg := 0 ;
   	AlarmAnalog[22].EnableCfg := 0 ;
   END_IF;
   AnalogPoint[22].Address := 22 ;
   AnalogPoint[22].RawMin := 5529 ;
   AnalogPoint[22].RawMax := 27648 ;
   AnalogPoint[22].RealCfg := 1 ;
   AnalogPoint[22].OverrideCfg := 1 ;
   AlarmAnalog[22].FeedPumpEnable := 0 ;
   AlarmAnalog[22].FeedPumpTag := 0 ;
   AlarmAnalog[22].TransferPumpEnable := 0 ;
   AlarmAnalog[22].TransferPumpTag := 0 ;
   AlarmAnalog[22].Disable := 0 ;
   AlarmAnalog[22].HIHIEnable := 0 ;
   
   (*Reset Loop : Set to 0 the AnalogPoint[23 to 27].EnableCfg
   ============================================================*)
   FOR Config.IndexAP := 23 to 27 by 1 do
   	AnalogPoint[Config.IndexAP].EnableCfg := 0 ;
   	AlarmAnalog[Config.IndexAP].EnableCfg := 0 ;
   End_for ;
   
   (*AnalogPoint[28]: Exchange AI#1
   ============================================================*)
   (*Set to 1 to use this AnalogPoint*)
   If Options.External_IO then
   	AnalogPoint[28].EnableCfg := 1 ;
   	AlarmAnalog[28].EnableCfg := 1 ;
   else
   	AnalogPoint[28].EnableCfg := 0 ;
   	AlarmAnalog[28].EnableCfg := 0 ;
   End_if ;
   (*Default Configuration *)
   AnalogPoint[28].Address := 28 ;
   AnalogPoint[28].RawMin := 6553 ;
   AnalogPoint[28].RawMax := 32767 ;
   AnalogPoint[28].RealCfg := 1 ;
   AnalogPoint[28].OverrideCfg := 1 ;
   AlarmAnalog[28].FeedPumpEnable := 0 ;
   AlarmAnalog[28].FeedPumpTag := 0 ;
   AlarmAnalog[28].TransferPumpEnable := 0 ;
   AlarmAnalog[28].TransferPumpTag := 0 ;
   AlarmAnalog[28].Disable := 0 ;
   AlarmAnalog[28].HIHIEnable := 0 ;
   
   (*AnalogPoint[29]: Exchange AI#2
   ============================================================*)
   (*Set to 1 to use this AnalogPoint*)
   If Options.External_IO then
   	AnalogPoint[29].EnableCfg := 1 ;
   	AlarmAnalog[29].EnableCfg := 1 ;
   else
   	AnalogPoint[29].EnableCfg := 0 ;
   	AlarmAnalog[29].EnableCfg := 0 ;
   End_if ;
   (*Default Configuration *)
   AnalogPoint[29].Address := 29 ;
   AnalogPoint[29].RawMin := 6553 ;
   AnalogPoint[29].RawMax := 32767 ;
   AnalogPoint[29].RealCfg := 1 ;
   AnalogPoint[29].OverrideCfg := 1 ;
   AlarmAnalog[29].FeedPumpEnable := 0 ;
   AlarmAnalog[29].FeedPumpTag := 0 ;
   AlarmAnalog[29].TransferPumpEnable := 0 ;
   AlarmAnalog[29].TransferPumpTag := 0 ;
   AlarmAnalog[29].Disable := 0 ;
   AlarmAnalog[29].HIHIEnable := 0 ;
   
   (*AnalogPoint[30]: Exchange AI#3
   ============================================================*)
   (*Set to 1 to use this AnalogPoint*)
   If Options.External_IO then
   	AnalogPoint[30].EnableCfg := 1 ;
   	AlarmAnalog[30].EnableCfg := 1 ;
   else
   	AnalogPoint[30].EnableCfg := 0 ;
   	AlarmAnalog[30].EnableCfg := 0 ;
   End_if ;
   (*Default Configuration *)
   AnalogPoint[30].Address := 30 ;
   AnalogPoint[30].RawMin := 6553 ;
   AnalogPoint[30].RawMax := 32767 ;
   AnalogPoint[30].RealCfg := 1 ;
   AnalogPoint[30].OverrideCfg := 1 ;
   AlarmAnalog[30].FeedPumpEnable := 0 ;
   AlarmAnalog[30].FeedPumpTag := 0 ;
   AlarmAnalog[30].TransferPumpEnable := 0 ;
   AlarmAnalog[30].TransferPumpTag := 0 ;
   AlarmAnalog[30].Disable := 0 ;
   AlarmAnalog[30].HIHIEnable := 0 ;
   
   (*AnalogPoint[31]: Exchange AI#4
   ============================================================*)
   (*Set to 1 to use this AnalogPoint*)
   If Options.External_IO then
   	AnalogPoint[31].EnableCfg := 1 ;
   	AlarmAnalog[31].EnableCfg := 1 ;
   else
   	AnalogPoint[31].EnableCfg := 0 ;
   	AlarmAnalog[31].EnableCfg := 0 ;
   End_if ;
   (*Default Configuration *)
   AnalogPoint[31].Address := 31 ;
   AnalogPoint[31].RawMin := 6553 ;
   AnalogPoint[31].RawMax := 32767 ;
   AnalogPoint[31].RealCfg := 1 ;
   AnalogPoint[31].OverrideCfg := 1 ;
   AlarmAnalog[31].FeedPumpEnable := 0 ;
   AlarmAnalog[31].FeedPumpTag := 0 ;
   AlarmAnalog[31].TransferPumpEnable := 0 ;
   AlarmAnalog[31].TransferPumpTag := 0 ;
   AlarmAnalog[31].Disable := 0 ;
   AlarmAnalog[31].HIHIEnable := 0 ;
   
   (*Reset Loop : Set to 0 the AnalogPoint[32 to 39].EnableCfg
   ============================================================*)
   FOR Config.IndexAP := 32 to 39 by 1 do
   	AnalogPoint[Config.IndexAP].EnableCfg := 0 ;
   	AlarmAnalog[Config.IndexAP].EnableCfg := 0 ;
   End_for ;
   
   (*AnalogPoint[40]: Differential Pressure DP
   ============================================================*)
   AnalogPoint[40].EnableCfg := 1 ;
   AnalogPoint[40].Address := 40 ;
   AnalogPoint[40].RawMin := 6553 ;
   AnalogPoint[40].RawMax := 32767 ;
   AnalogPoint[40].RealCfg := 0 ;
   AnalogPoint[40].OverrideCfg := 1 ;
   AlarmAnalog[40].FeedPumpEnable := 1 ;
   AlarmAnalog[40].FeedPumpTag := 1 ;
   AlarmAnalog[40].TransferPumpEnable := 0 ;
   AlarmAnalog[40].TransferPumpTag := 0 ;
   AlarmAnalog[40].EnableCfg := 1 ;
   AlarmAnalog[40].Disable := 0 ;
   AlarmAnalog[40].HIHIEnable := 0 ;
   
   (*AnalogPoint[41]: Trans-Membrane Pressure TMP
   ============================================================*)
   AnalogPoint[41].EnableCfg := 1 ;
   AnalogPoint[41].Address := 41 ;
   AnalogPoint[41].RawMin := 6553 ;
   AnalogPoint[41].RawMax := 32767 ;
   AnalogPoint[41].RealCfg := 0 ;
   AnalogPoint[41].OverrideCfg := 1 ;
   AlarmAnalog[41].FeedPumpEnable := 1 ;
   AlarmAnalog[41].FeedPumpTag := 1 ;
   AlarmAnalog[41].TransferPumpEnable := 0 ;
   AlarmAnalog[41].TransferPumpTag := 0 ;
   AlarmAnalog[41].EnableCfg := 1 ;
   AlarmAnalog[41].Disable := 0 ;
   AlarmAnalog[41].HIHIEnable := 0 ;
   
   (*AnalogPoint[42]: Feed Flow FI003
   ============================================================*)
   AnalogPoint[42].EnableCfg := 1 ;
   AnalogPoint[42].Address := 42 ;
   AnalogPoint[42].RawMin := 6553 ;
   AnalogPoint[42].RawMax := 32767 ;
   AnalogPoint[42].RealCfg := 0 ;
   AnalogPoint[42].OverrideCfg := 1 ;
   AlarmAnalog[42].FeedPumpEnable := 1 ;
   AlarmAnalog[42].FeedPumpTag := 1 ;
   AlarmAnalog[42].TransferPumpEnable := 0 ;
   AlarmAnalog[42].TransferPumpTag := 0 ;
   AlarmAnalog[42].EnableCfg := 1 ;
   AlarmAnalog[42].Disable := 0 ;
   AlarmAnalog[42].HIHIEnable := 0 ;
   
   (*AnalogPoint[43]: Spare
   ============================================================*)
   AnalogPoint[43].EnableCfg := 0 ;
   AnalogPoint[43].Address := 43 ;
   AnalogPoint[43].RawMin := 6553 ;
   AnalogPoint[43].RawMax := 32767 ;
   AnalogPoint[43].RealCfg := 0 ;
   AnalogPoint[43].OverrideCfg := 1 ;
   AlarmAnalog[43].FeedPumpEnable := 0 ;
   AlarmAnalog[43].FeedPumpTag := 0 ;
   AlarmAnalog[43].TransferPumpEnable := 0 ;
   AlarmAnalog[43].TransferPumpTag := 0 ;
   AlarmAnalog[43].EnableCfg := 0 ;
   AlarmAnalog[43].Disable := 0 ;
   AlarmAnalog[43].HIHIEnable := 0 ;
   
   (*AnalogPoint[44]: Feed Tank Volume LI101
   ============================================================*)
   AnalogPoint[44].EnableCfg := 1 ;
   AnalogPoint[44].Address := 44 ;
   AnalogPoint[44].RawMin := 6553 ;
   AnalogPoint[44].RawMax := 32767 ;
   AnalogPoint[44].RealCfg := 0 ;
   AnalogPoint[44].OverrideCfg := 1 ;
   AlarmAnalog[44].FeedPumpEnable := 1 ;
   AlarmAnalog[44].FeedPumpTag := 1 ;
   AlarmAnalog[44].TransferPumpEnable := 0 ;
   AlarmAnalog[44].TransferPumpTag := 0 ;
   AlarmAnalog[44].EnableCfg := 1 ;
   AlarmAnalog[44].Disable := 0 ;
   AlarmAnalog[44].HIHIDisable := NOT SIC002.RunStatus ;
   AlarmAnalog[44].HIDisable := NOT SIC002.RunStatus ;
   AlarmAnalog[44].HIHIEnable := 0 ;
   
   (*AnalogPoint[45]: Normalized Water Permeability NWP
   ============================================================*)
   AnalogPoint[45].EnableCfg := 1 ;
   AnalogPoint[45].Address := 45 ;
   AnalogPoint[45].RawMin := 6553 ;
   AnalogPoint[45].RawMax := 32767 ;
   AnalogPoint[45].RealCfg := 0 ;
   AnalogPoint[45].OverrideCfg := 0 ;
   AlarmAnalog[45].FeedPumpEnable := 0 ;
   AlarmAnalog[45].FeedPumpTag := 0 ;
   AlarmAnalog[45].TransferPumpEnable := 0 ;
   AlarmAnalog[45].TransferPumpTag := 0 ;
   AlarmAnalog[45].EnableCfg := 0 ;
   AlarmAnalog[45].Disable := 0 ;
   AlarmAnalog[45].HIHIEnable := 0 ;
   
   (*AnalogPoint[46]: Membrane Permeability PERM
   ============================================================*)
   AnalogPoint[46].EnableCfg := 1 ;
   AnalogPoint[46].Address := 46 ;
   AnalogPoint[46].RawMin := 6553 ;
   AnalogPoint[46].RawMax := 32767 ;
   AnalogPoint[46].RealCfg := 0 ;
   AnalogPoint[46].OverrideCfg := 0 ;
   AlarmAnalog[46].FeedPumpEnable := 0 ;
   AlarmAnalog[46].FeedPumpTag := 0 ;
   AlarmAnalog[46].TransferPumpEnable := 0 ;
   AlarmAnalog[46].TransferPumpTag := 0 ;
   AlarmAnalog[46].EnableCfg := 0 ;
   AlarmAnalog[46].Disable := 0 ;
   AlarmAnalog[46].HIHIEnable := 0 ;
   
   (*Reset Loop : Set to 0 the AnalogPoint[47 to 49].EnableCfg
   ============================================================*)
   FOR Config.IndexAP := 47 to 49 by 1 do
   	AnalogPoint[Config.IndexAP].EnableCfg := 0 ;
   	AlarmAnalog[Config.IndexAP].EnableCfg := 0 ;
   End_for ;
   
END_ROUTINE

ROUTINE Config_ControlLoop   (* structured text *)
   (* =======================================================================
   	Config ControlLoop : Configure ControlLoop Structure
   
   	List of treatments
   		- ControlLoop[1] : FIC003 Feed Pump Control Loop
   		- ControlLoop[2] : LIC101 Level Control Loop
   		- ControlLoop[3] : PCV101 Retentate Control Valve Control Loop
   		- ControlLoop[4] : PCV101 Retentate Control Valve Control Loop 5ms
   		- ControlLoop[5] : PCV201 Filtrate Control Valve Control Loop
   		- ControlLoop[6] : PCV201 Filtrate Control Valve Control Loop 5ms
   		- ControlLoop[7] : TIC101 TCU Temperature Control Loop
   		- Reset Loop : Disable unused ControlLoop and Deviation Alarm
   
   -----------------------------------------------------------------------------------------------------------------------------------------------------
   	History
   		2019-DEC-24 - Merck - Q. Spindler - Initial version for Candidate Release 1.00.00.00.a
   		2021-APR-19 - Merck - Q. Spindler - Modifications for Candidate Release 1.00.00.00.e
                       - Change PCV Full Open/Close timer from 1sec to 3sec
   					- Change TIC101 Range max to 50
   		2022-SEP-22 - Actemium - J. Jaekel - Modifications for Candidate Release 1.01.00.01.a
   					- Add ExternalTCU option to TIC101 ControlLoop
   =========================================================================*)
   
   (* FIC003 Feed Pump Control Loop
   =========================================================================*)
   (*Index set with ControlLoop number*)
   Config.IndexCL := 1 ;
   (*ControlLoop data structure configuration*)
   ControlLoop[1].LoopCfg := 1 ;
   ControlLoop[1].Auto4 := 0;
   ControlLoop[1].RampEnable := 1;
   ControlLoop[1].PIDEnable := 1;
   ControlLoop[1].StepIncrement := 0;
   ControlLoop[1].CycleTime := 0;
   ControlLoop[1].SPAuto4 := 0;
   ControlLoop[1].RangeMin := 0;
   ControlLoop[1].RangeMax := 100;
   ControlLoop[1].RampTimer.PRE := 3600000;
   ControlLoop[1].PIDTimer.PRE := 250;
   ControlLoop[1].CycleTimer.PRE := 2000;
   ControlLoop[1].DigitalOutput := 0;
   ControlLoop[1].RampCfg := 0;
   ControlLoop[1].Auto1Cfg := 1;
   ControlLoop[1].Auto2Cfg := 1;
   ControlLoop[1].Auto3Cfg := 1;
   ControlLoop[1].Auto4Cfg := 0;
   ControlLoop[1].Auto1PVCfg := 42; //FI003
   ControlLoop[1].Auto2PVCfg := 40; //DP
   ControlLoop[1].Auto3PVCfg := 5; //PI001
   ControlLoop[1].Auto4PVCfg := 0;
   ControlLoop[1].Auto1RangeMax := FI003.ScaledMax;
   ControlLoop[1].Auto2RangeMax := DP.ScaledMax;
   ControlLoop[1].Auto3RangeMax := PI001.ScaledMax;
   ControlLoop[1].Auto4RangeMax := 0;
   ControlLoop[1].AutoSwitchEnable := 0;
   ControlLoop[1].OutputAddress := 2;
   (*Deviation data structure configuration*)
   AlarmDeviation[1].EnableCfg := 1;
   
   (* LIC101 Level Control Loop
   =========================================================================*)
   (*ControlLoop data structure configuration*)
   IF Options.TransferFlow THEN
   	ControlLoop[2].Auto2Cfg := 1;
   ELSE
   	ControlLoop[2].Auto2Cfg := 0;
   	ControlLoop[2].Auto2 := 0;
   	ControlLoop[2].SPAuto2 := 0;
   END_IF;
   ControlLoop[2].LoopCfg := 1 ;
   ControlLoop[2].Auto3 := 0;
   ControlLoop[2].Auto4 := 0;
   ControlLoop[2].RampEnable := 1;
   ControlLoop[2].PIDEnable := 1;
   ControlLoop[2].StepIncrement := 0;
   ControlLoop[2].CycleTime := 0;
   ControlLoop[2].SPAuto3 := 0;
   ControlLoop[2].SPAuto4 := 0;
   ControlLoop[2].RangeMin := 0;
   ControlLoop[2].RangeMax := 100;
   ControlLoop[2].RampTimer.PRE := 3600000;
   ControlLoop[2].PIDTimer.PRE := 250;
   ControlLoop[2].CycleTimer.PRE := 2000;
   ControlLoop[2].DigitalOutput := 0;
   ControlLoop[2].RampCfg := 0;
   ControlLoop[2].Auto1Cfg := 1;
   ControlLoop[2].Auto3Cfg := 0;
   ControlLoop[2].Auto4Cfg := 0;
   ControlLoop[2].Auto1PVCfg := 44; //LI101
   ControlLoop[2].Auto2PVCfg := 20; //FI401
   ControlLoop[2].Auto3PVCfg := 0;
   ControlLoop[2].Auto4PVCfg := 0;
   ControlLoop[2].Auto1RangeMax := LI101.ScaledMax;
   ControlLoop[2].Auto2RangeMax := FI401.ScaledMax;
   ControlLoop[2].Auto3RangeMax := 0;
   ControlLoop[2].Auto4RangeMax := 0;
   ControlLoop[2].AutoSwitchEnable := 0;
   ControlLoop[2].OutputAddress := 1;
   (*Deviation data structure configuration*)
   AlarmDeviation[2].EnableCfg := 1;
   
   (* PCV101 Retentate Control Valve Control Loop
   =========================================================================*)
   (*ControlLoop data structure configuration*)
   ControlLoop[3].LoopCfg := 1 ;
   ControlLoop[3].Auto3 := 0;
   ControlLoop[3].Auto4 := 0;
   ControlLoop[3].PIDEnable := 1;
   ControlLoop[3].StepIncrement := 0;
   ControlLoop[3].CycleTime := 0;
   ControlLoop[3].SPAuto3 := 0;
   ControlLoop[3].SPAuto4 := 0;
   ControlLoop[3].RangeMin := 0;
   ControlLoop[3].RangeMax := 100;
   ControlLoop[3].RampTimer.PRE := 3600000;
   ControlLoop[3].PIDTimer.PRE := 250;
   ControlLoop[3].CycleTimer.PRE := 2000;
   ControlLoop[3].On := 0;
   ControlLoop[3].DigitalOutput := 0;
   ControlLoop[3].RampCfg := 0;
   ControlLoop[3].Auto1Cfg := 1;
   ControlLoop[3].Auto2Cfg := 1;
   ControlLoop[3].Auto3Cfg := 0;
   ControlLoop[3].Auto4Cfg := 0;
   ControlLoop[3].Auto1PVCfg := 6; //PI101
   ControlLoop[3].Auto2PVCfg := 41; //TMP
   ControlLoop[3].Auto3PVCfg := 0;
   ControlLoop[3].Auto4PVCfg := 0;
   ControlLoop[3].Auto1RangeMax := PI101.ScaledMax;
   ControlLoop[3].Auto2RangeMax := TMP.ScaledMax;
   ControlLoop[3].Auto3RangeMax := 0;
   ControlLoop[3].Auto4RangeMax := 0;
   ControlLoop[3].AutoSwitchEnable := 0;
   ControlLoop[3].OutputAddress := 3;
   (*Deviation data structure configuration*)
   AlarmDeviation[3].EnableCfg := 1;
   (*PCV Control : 0-100 %Clo*)
   PCV101_Control.FullOpenSP := 0 ;
   PCV101_Control.FullCloseSP := 100 ;
   PCV101_Control.FullOpenResetTimer.PRE := 3000 ;
   PCV101_Control.FullCloseResetTimer.PRE := 3000 ;
   
   (* PCV101 Retentate Control Valve Control Loop 5ms
   =========================================================================*)
   (*ControlLoop data structure configuration*)
   ControlLoop[4].LoopCfg := 0 ;
   ControlLoop[4].Manual := 0;
   ControlLoop[4].Auto1 := 0;
   ControlLoop[4].Auto2 := 0;
   ControlLoop[4].Auto3 := 0;
   ControlLoop[4].Auto4 := 0;
   ControlLoop[4].PIDEnable := 1;
   ControlLoop[4].RampEnable := 0;
   ControlLoop[4].StepIncrement := 0;
   ControlLoop[4].CycleTime := 0;
   ControlLoop[4].SPAuto1 := 0;
   ControlLoop[4].SPAuto2 := 0;
   ControlLoop[4].SPAuto3 := 0;
   ControlLoop[4].SPAuto4 := 0;
   ControlLoop[4].RangeMin := 0;
   ControlLoop[4].RangeMax := 100;
   ControlLoop[4].RampTimer.PRE := 3600000;
   ControlLoop[4].PIDTimer.PRE := 250;
   ControlLoop[4].CycleTimer.PRE := 2000;
   ControlLoop[4].On := 0;
   ControlLoop[4].DigitalOutput := 0;
   ControlLoop[4].RampCfg := 0;
   ControlLoop[4].Auto1Cfg := 0;
   ControlLoop[4].Auto2Cfg := 0;
   ControlLoop[4].Auto3Cfg := 0;
   ControlLoop[4].Auto4Cfg := 0;
   ControlLoop[4].Auto1PVCfg := 0;
   ControlLoop[4].Auto2PVCfg := 0;
   ControlLoop[4].Auto3PVCfg := 0;
   ControlLoop[4].Auto4PVCfg := 0;
   ControlLoop[4].Auto1RangeMax := 0;
   ControlLoop[4].Auto2RangeMax := 0;
   ControlLoop[4].Auto3RangeMax := 0;
   ControlLoop[4].Auto4RangeMax := 0;
   ControlLoop[4].AutoSwitchEnable := 0;
   ControlLoop[4].OutputAddress := 3;
   ControlLoop[4].PID.KP := 0.2;
   ControlLoop[4].PID.KD := 0.01;
   ControlLoop[4].PID.DB := 0.3;
   ControlLoop[4].PID.UPD := 0.005;
   ControlLoop[4].PID.MAXS := 100;
   ControlLoop[4].PID.MAXO := 100;
   ControlLoop[4].PID.MAXI := 100;
   ControlLoop[4].PID.MAXCV := 100;
   ControlLoop[4].PID.MAXTIE := 4095;
   
   (* PCV201 Filtrate Control Valve Control Loop
   =========================================================================*)
   (*ControlLoop data structure configuration*)
   ControlLoop[5].LoopCfg := 1 ;
   ControlLoop[5].Auto3 := 0;
   ControlLoop[5].Auto4 := 0;
   ControlLoop[5].PIDEnable := 1;
   ControlLoop[5].StepIncrement := 0;
   ControlLoop[5].CycleTime := 0;
   ControlLoop[5].SPAuto3 := 0;
   ControlLoop[5].SPAuto4 := 0;
   ControlLoop[5].RangeMin := 0;
   ControlLoop[5].RangeMax := 100;
   ControlLoop[5].RampTimer.PRE := 3600000;
   ControlLoop[5].PIDTimer.PRE := 250;
   ControlLoop[5].CycleTimer.PRE := 2000;
   ControlLoop[5].On := 0;
   ControlLoop[5].DigitalOutput := 0;
   ControlLoop[5].RampCfg := 0;
   ControlLoop[5].Auto1Cfg := 1;
   ControlLoop[5].Auto2Cfg := 1;
   ControlLoop[5].Auto3Cfg := 0;
   ControlLoop[5].Auto4Cfg := 0;
   ControlLoop[5].Auto1PVCfg := 2; // FI201
   ControlLoop[5].Auto2PVCfg := 41; // TMP
   ControlLoop[5].Auto3PVCfg := 0;
   ControlLoop[5].Auto4PVCfg := 0;
   ControlLoop[5].Auto1RangeMax := FI201.ScaledMax;
   ControlLoop[5].Auto2RangeMax := TMP.ScaledMax;
   ControlLoop[5].Auto3RangeMax := 0;
   ControlLoop[5].Auto4RangeMax := 0;
   ControlLoop[5].AutoSwitchEnable := 0;
   ControlLoop[5].OutputAddress := 4;
   (*Deviation data structure configuration*)
   AlarmDeviation[5].EnableCfg := 1;
   (*PCV Control : 0-100 %opn*)
   PCV201_Control.FullOpenSP := 100 ;
   PCV201_Control.FullCloseSP := 0 ;
   PCV201_Control.FullOpenResetTimer.PRE := 3000 ;
   PCV201_Control.FullCloseResetTimer.PRE := 3000 ;
   
   
   (* PCV201 Filtrate Control Valve Control Loop
   =========================================================================*)
   
   (*ControlLoop data structure configuration*)
   ControlLoop[6].LoopCfg := 0 ;
   ControlLoop[6].Manual := 0;
   ControlLoop[6].Auto1 := 0;
   ControlLoop[6].Auto2 := 0;
   ControlLoop[6].Auto3 := 0;
   ControlLoop[6].Auto4 := 0;
   ControlLoop[6].PIDEnable := 1;
   ControlLoop[6].RampEnable := 0;
   ControlLoop[6].StepIncrement := 0;
   ControlLoop[6].CycleTime := 0;
   ControlLoop[6].SPAuto1 := 0;
   ControlLoop[6].SPAuto2 := 0;
   ControlLoop[6].SPAuto3 := 0;
   ControlLoop[6].SPAuto4 := 0;
   ControlLoop[6].RangeMin := 0;
   ControlLoop[6].RangeMax := 100;
   ControlLoop[6].RampTimer.PRE := 3600000;
   ControlLoop[6].PIDTimer.PRE := 250;
   ControlLoop[6].CycleTimer.PRE := 2000;
   ControlLoop[6].On := 0;
   ControlLoop[6].DigitalOutput := 0;
   ControlLoop[6].RampCfg := 0;
   ControlLoop[6].Auto1Cfg := 0;
   ControlLoop[6].Auto2Cfg := 0;
   ControlLoop[6].Auto3Cfg := 0;
   ControlLoop[6].Auto4Cfg := 0;
   ControlLoop[6].Auto1PVCfg := 0;
   ControlLoop[6].Auto2PVCfg := 0;
   ControlLoop[6].Auto3PVCfg := 0;
   ControlLoop[6].Auto4PVCfg := 0;
   ControlLoop[6].Auto1RangeMax := 0;
   ControlLoop[6].Auto2RangeMax := 0;
   ControlLoop[6].Auto3RangeMax := 0;
   ControlLoop[6].Auto4RangeMax := 0;
   ControlLoop[6].AutoSwitchEnable := 0;
   ControlLoop[6].OutputAddress := 4;
   ControlLoop[6].PID.KP := 0.3;
   ControlLoop[6].PID.KD := 0.01;
   ControlLoop[6].PID.DB := 0.3;
   ControlLoop[6].PID.UPD := 0.005;
   ControlLoop[6].PID.MAXS := 100;
   ControlLoop[6].PID.MAXO := 100;
   ControlLoop[6].PID.MAXI := 100;
   ControlLoop[6].PID.MAXCV := 100;
   ControlLoop[6].PID.MAXTIE := 4095;
   
   (* TIC101 TCU Temperature Control Loop
   =========================================================================*)
   (*ControlLoop data structure configuration*)
   IF Options.FeedTank and ExternalTCU THEN
   	ControlLoop[7].LoopCfg := 1;
   	AlarmDeviation[7].EnableCfg := 1;
   ELSE
   	ControlLoop[7].LoopCfg := 0;
   	AlarmDeviation[7].EnableCfg := 0;
   END_IF;
   ControlLoop[7].Auto2 := 0;
   ControlLoop[7].Auto3 := 0;
   ControlLoop[7].Auto4 := 0;
   ControlLoop[7].RampEnable := 0;
   ControlLoop[7].PIDEnable := 1;
   ControlLoop[7].StepIncrement := 0;
   ControlLoop[7].CycleTime := 0;
   ControlLoop[7].SPAuto2 := 0;
   ControlLoop[7].SPAuto3 := 0;
   ControlLoop[7].SPAuto4 := 0;
   ControlLoop[7].RangeMin := 0;
   ControlLoop[7].RangeMax := 50;
   ControlLoop[7].RampTimer.PRE := 3600000;
   ControlLoop[7].PIDTimer.PRE := 250;
   ControlLoop[7].CycleTimer.PRE := 2000;
   ControlLoop[7].DigitalOutput := 0;
   ControlLoop[7].RampCfg := 0;
   ControlLoop[7].Auto1Cfg := 1;
   ControlLoop[7].Auto2Cfg := 0;
   ControlLoop[7].Auto3Cfg := 0;
   ControlLoop[7].Auto4Cfg := 0;
   ControlLoop[7].Auto1PVCfg := 13; //TI101
   ControlLoop[7].Auto2PVCfg := 0;
   ControlLoop[7].Auto3PVCfg := 0;
   ControlLoop[7].Auto4PVCfg := 0;
   ControlLoop[7].Auto1RangeMax := TI101.ScaledMax;
   ControlLoop[7].Auto2RangeMax := 0;
   ControlLoop[7].Auto3RangeMax := 0;
   ControlLoop[7].Auto4RangeMax := 0;
   ControlLoop[7].AutoSwitchEnable := 0;
   ControlLoop[7].OutputAddress := 6; // TCU101_AO
   
   (*Reset Loop : Disable unused ControlLoop and Deviation Alarm
   ============================================================*)
   ControlLoop[0].LoopCfg := 0 ;
   AlarmDeviation[0].EnableCfg := 0;
   AlarmDeviation[0].Override := 1;
   AlarmDeviation[0].Disable := 1;
   ControlLoop[4].LoopCfg := 0 ;
   AlarmDeviation[4].EnableCfg := 0;
   AlarmDeviation[4].Override := 1;
   AlarmDeviation[4].Disable := 1;
   ControlLoop[6].LoopCfg := 0 ;
   AlarmDeviation[6].EnableCfg := 0;
   AlarmDeviation[6].Override := 1;
   AlarmDeviation[6].Disable := 1;
   
   FOR Config.IndexCL := 8 to 19 do
   	ControlLoop[Config.IndexCL].LoopCfg := 0 ;
   	AlarmDeviation[Config.IndexCL].EnableCfg := 0;
   	AlarmDeviation[Config.IndexCL].Override := 1;
   	AlarmDeviation[Config.IndexCL].Disable := 1;
   End_for ;
END_ROUTINE
